// TIA Portal V20 export
// export: Created 2026-10-20T12:47:21.9915101Z, ExportSetting WithDefaults, DisplayName Totally Integrated Automation Portal, DisplayVersion V20 Update 6, DisplayName TIA Portal Openness, DisplayVersion V20 Update 6, DisplayName TIA Portal Version Control Interface, DisplayVersion V20 Update 6, DisplayName SINAMICS Startdrive Advanced, DisplayVersion V20 SP1, DisplayName SINAMICS Startdrive G130, G150, S120, S150, SINAMICS MV, G220, S200, S210, DisplayVersion V20 SP1, DisplayName SINAMICS Startdrive G110M, G120, G120C, G120D, G120P, G115D, DisplayVersion V20 SP1, DisplayName STEP 7 Professional, DisplayVersion V20 Update 6, DisplayName STEP 7 Safety, DisplayVersion V20 Update 2, DisplayName WinCC Basic/Comfort/Advanced, DisplayVersion V20 Update 6, DisplayName WinCC Unified, DisplayVersion V20 Update 6
FUNCTION "INPUTS" : Void   // FC25, SCL
{ S7_Optimized_Access := 'TRUE' }
VERSION : 0.1
// stored: AutoNumber true, IsIECCheckEnabled false, SetENOAutomatically false, UDAEnableTagReadback false
BEGIN
   REGION SYSTEM 1
       REGION EXTRACTOR CONVEYOR
           "Control_DB".ECnv_Sys[1].Inputs.Left := "CVTD1 SENSOR CONVEYOR LEFT";
           "Control_DB".ECnv_Sys[1].Inputs.Lpd1 := "CVTD1 SENSOR CONVEYOR LEFT (PALLET DETECT 1)";
           "Control_DB".ECnv_Sys[1].Inputs.Center := "CVTD1 SENSOR CONVEYOR CENTER";
           "Control_DB".ECnv_Sys[1].Inputs.Right := "CVTD1 SENSOR CONVEYOR RIGHT";
           "Control_DB".ECnv_Sys[1].Inputs.Rpd1 := "CVTD1 SENSOR CONVEYOR RIGHT (PALLET DETECT 1)";

           "T_OH_Left_1".TOF(IN := "CVTD1 OVERHANG LEFT" OR NOT "Control_DB".VTD_Sys[1].Running,
                             PT := T#200ms);
           "Control_DB".ECnv_Sys[1].Inputs.Overhang_Left := "T_OH_Left_1".Q;

           "T_OH_Right_1".TOF(IN := "CVTD1 OVERHANG RIGHT" OR NOT "Control_DB".VTD_Sys[1].Running,
                              PT := T#200ms);
           "Control_DB".ECnv_Sys[1].Inputs.Overhang_Right := "T_OH_Right_1".Q;

           "Control_DB".ECnv_Sys[1].Inputs.VFD_Status := "CVTD1_StatusWord";
           "Control_DB".ECnv_Sys[1].Inputs.VFD_ActualCurrent := WORD_TO_INT("CVTD1_ActualCurrent");
           "Control_DB".ECnv_Sys[1].Inputs.VFD_Speed_Actual := WORD_TO_INT("CVTD1_ActualSpeed");
           "Control_DB".ECnv_Sys[1].Inputs.VFD_ActualTorque := WORD_TO_INT("CVTD1_ActualTorque");
       END_REGION

       REGION BUFFER CONVEYORS
           REGION LEVEL 1
               //BUFFER CONVEYOR LEVEL 1 - CONVEYOR 1
               "Control_DB".LCnv_Sys[1].Cnv_Level[1].Cnv1.Inputs.Left := NOT "C1101 - SENSOR CNV LEFT";
               "Control_DB".LCnv_Sys[1].Cnv_Level[1].Cnv1.Inputs.Lpd1 := NOT "C1101 - SENSOR CNV LEFT (PALLET DETECT 1)";
               "Control_DB".LCnv_Sys[1].Cnv_Level[1].Cnv1.Inputs.Lpd2 := "C1101 - SENSOR CNV LEFT (PALLET DETECT 2)";
               "Control_DB".LCnv_Sys[1].Cnv_Level[1].Cnv1.Inputs.Right := NOT "C1101 - SENSOR CNV RIGHT";
               "Control_DB".LCnv_Sys[1].Cnv_Level[1].Cnv1.Inputs.Rpd1 := NOT "C1101 - SENSOR CNV RIGHT (PALLET DETECT 1)";
               "Control_DB".LCnv_Sys[1].Cnv_Level[1].Cnv1.Inputs.Rpd2 := NOT "C1101 - SENSOR CNV RIGHT (PALLET DETECT 2)";
               "Control_DB".LCnv_Sys[1].Cnv_Level[1].Cnv1.Inputs.Sdetect1 := NOT "C1101 - SHUTTLE IN POSITION 1";
               "Control_DB".LCnv_Sys[1].Cnv_Level[1].Cnv1.Inputs.Sdetect2 := NOT "C1101 - SHUTTLE IN POSITION 2";

               "Control_DB".LCnv_Sys[1].Cnv_Level[1].Cnv1.Inputs.VFD_Status := "C1101_StatusWord";
               "Control_DB".LCnv_Sys[1].Cnv_Level[1].Cnv1.Inputs.VFD_ActualCurrent := WORD_TO_INT("C1101_ActualCurrent");
               "Control_DB".LCnv_Sys[1].Cnv_Level[1].Cnv1.Inputs.VFD_Speed_Actual := WORD_TO_INT("C1101_ActualSpeed");
               "Control_DB".LCnv_Sys[1].Cnv_Level[1].Cnv1.Inputs.VFD_ActualTorque := WORD_TO_INT("C1101_ActualTorque");

               //BUFFER CONVEYOR LEVEL 1 - CONVEYOR 2
               "Control_DB".LCnv_Sys[1].Cnv_Level[1].Cnv2.Inputs.Left := NOT "C1201 - SENSOR CNV LEFT";
               "Control_DB".LCnv_Sys[1].Cnv_Level[1].Cnv2.Inputs.Lpd1 := NOT "C1201 - SENSOR CNV LEFT (PALLET DETECT 1)";
               "Control_DB".LCnv_Sys[1].Cnv_Level[1].Cnv2.Inputs.Lpd2 := NOT "C1201 - SENSOR CNV LEFT (PALLET DETECT 2)";
               "Control_DB".LCnv_Sys[1].Cnv_Level[1].Cnv2.Inputs.Right := NOT "C1201 - SENSOR CNV RIGHT";
               "Control_DB".LCnv_Sys[1].Cnv_Level[1].Cnv2.Inputs.Rpd1 := NOT "C1201 - SENSOR CNV RIGHT (PALLET DETECT 1)";
               "Control_DB".LCnv_Sys[1].Cnv_Level[1].Cnv2.Inputs.Rpd2 := NOT "C1201 - SENSOR CNV RIGHT (PALLET DETECT 2)";
               "Control_DB".LCnv_Sys[1].Cnv_Level[1].Cnv2.Inputs.Sdetect1 := NOT "C1201 - SHUTTLE IN POSITION 1";
               "Control_DB".LCnv_Sys[1].Cnv_Level[1].Cnv2.Inputs.Sdetect2 := NOT "C1201 - SHUTTLE IN POSITION 2";

               "Control_DB".LCnv_Sys[1].Cnv_Level[1].Cnv2.Inputs.VFD_Status := "C1201_StatusWord";
               "Control_DB".LCnv_Sys[1].Cnv_Level[1].Cnv2.Inputs.VFD_ActualCurrent := WORD_TO_INT("C1201_ActualCurrent");
               "Control_DB".LCnv_Sys[1].Cnv_Level[1].Cnv2.Inputs.VFD_Speed_Actual := WORD_TO_INT("C1201_ActualSpeed");
               "Control_DB".LCnv_Sys[1].Cnv_Level[1].Cnv2.Inputs.VFD_ActualTorque := WORD_TO_INT("C1201_ActualTorque");
           END_REGION

           REGION LEVEL 2
               //BUFFER CONVEYOR LEVEL 2 - CONVEYOR 1
               "Control_DB".LCnv_Sys[1].Cnv_Level[2].Cnv1.Inputs.Left := NOT "C1102 - SENSOR CNV LEFT";
               "Control_DB".LCnv_Sys[1].Cnv_Level[2].Cnv1.Inputs.Lpd1 := NOT "C1102 - SENSOR CNV LEFT (PALLET DETECT 1)";
               "Control_DB".LCnv_Sys[1].Cnv_Level[2].Cnv1.Inputs.Lpd2 := NOT "C1102 - SENSOR CNV LEFT (PALLET DETECT 2)";
               "Control_DB".LCnv_Sys[1].Cnv_Level[2].Cnv1.Inputs.Right := NOT "C1102 - SENSOR CNV RIGHT";
               "Control_DB".LCnv_Sys[1].Cnv_Level[2].Cnv1.Inputs.Rpd1 := NOT "C1102 - SENSOR CNV RIGHT (PALLET DETECT 1)";
               "Control_DB".LCnv_Sys[1].Cnv_Level[2].Cnv1.Inputs.Rpd2 := NOT "C1102 - SENSOR CNV RIGHT (PALLET DETECT 2)";
               "Control_DB".LCnv_Sys[1].Cnv_Level[2].Cnv1.Inputs.Sdetect1 := NOT "C1102 - SHUTTLE IN POSITION 1";
               "Control_DB".LCnv_Sys[1].Cnv_Level[2].Cnv1.Inputs.Sdetect2 := NOT "C1102 - SHUTTLE IN POSITION 2";
               "Control_DB".LCnv_Sys[1].Cnv_Level[2].Cnv1.Safety_Stop_Cnrl.Inputs.DP_Extended := "C1102 - SENSOR SAFETY PIN1 UP";
               "Control_DB".LCnv_Sys[1].Cnv_Level[2].Cnv1.Safety_Stop_Cnrl.Inputs.DP_Retracted := "C1102 - SENSOR SAFETY PIN1 DOWN";

               IF "Shuttle_MQTT_DB".Shuttle_MQTT[3].Message.Shuttle_Status.Position_ID = "Settings_DB".LCnv_Sys[1].Cnv_Level[2].Cnv1.Barcode_ID THEN
                   "Control_DB".LCnv_Sys[1].Cnv_Level[2].Cnv1.Inputs.Shuttle_High := "Shuttle_MQTT_DB".Shuttle_MQTT[3].Message.Shuttle_Status.Sensor_Inputs.%X13;
               ELSIF "Shuttle_MQTT_DB".Shuttle_MQTT[4].Message.Shuttle_Status.Position_ID = "Settings_DB".LCnv_Sys[1].Cnv_Level[2].Cnv1.Barcode_ID THEN
                   "Control_DB".LCnv_Sys[1].Cnv_Level[2].Cnv1.Inputs.Shuttle_High := "Shuttle_MQTT_DB".Shuttle_MQTT[4].Message.Shuttle_Status.Sensor_Inputs.%X13;
               ELSIF "Shuttle_MQTT_DB".Shuttle_MQTT[5].Message.Shuttle_Status.Position_ID = "Settings_DB".LCnv_Sys[1].Cnv_Level[2].Cnv1.Barcode_ID THEN
                   "Control_DB".LCnv_Sys[1].Cnv_Level[2].Cnv1.Inputs.Shuttle_High := "Shuttle_MQTT_DB".Shuttle_MQTT[5].Message.Shuttle_Status.Sensor_Inputs.%X13;
               END_IF;

               "Control_DB".LCnv_Sys[1].Cnv_Level[2].Cnv1.Inputs.VFD_Status := "C1102_StatusWord";
               "Control_DB".LCnv_Sys[1].Cnv_Level[2].Cnv1.Inputs.VFD_ActualCurrent := WORD_TO_INT("C1102_ActualCurrent");
               "Control_DB".LCnv_Sys[1].Cnv_Level[2].Cnv1.Inputs.VFD_Speed_Actual := WORD_TO_INT("C1102_ActualSpeed");
               "Control_DB".LCnv_Sys[1].Cnv_Level[2].Cnv1.Inputs.VFD_ActualTorque := "C1102_ActualTorque";

               //BUFFER CONVEYOR LEVEL 2 - CONVEYOR 2
               "Control_DB".LCnv_Sys[1].Cnv_Level[2].Cnv2.Inputs.Left := NOT "C1202 - SENSOR CNV LEFT";
               "Control_DB".LCnv_Sys[1].Cnv_Level[2].Cnv2.Inputs.Lpd1 := NOT "C1202 - SENSOR CNV LEFT (PALLET DETECT 1)";
               "Control_DB".LCnv_Sys[1].Cnv_Level[2].Cnv2.Inputs.Lpd2 := NOT "C1202 - SENSOR CNV LEFT (PALLET DETECT 2)";
               "Control_DB".LCnv_Sys[1].Cnv_Level[2].Cnv2.Inputs.Right := NOT "C1202 - SENSOR CNV RIGHT";
               "Control_DB".LCnv_Sys[1].Cnv_Level[2].Cnv2.Inputs.Rpd1 := NOT "C1202 - SENSOR CNV RIGHT (PALLET DETECT 1)";
               "Control_DB".LCnv_Sys[1].Cnv_Level[2].Cnv2.Inputs.Rpd2 := NOT "C1202 - SENSOR CNV RIGHT (PALLET DETECT 2)";
               "Control_DB".LCnv_Sys[1].Cnv_Level[2].Cnv2.Inputs.Sdetect1 := NOT "C1202 - SHUTTLE IN POSITION 1";
               "Control_DB".LCnv_Sys[1].Cnv_Level[2].Cnv2.Inputs.Sdetect2 := NOT "C1202 - SHUTTLE IN POSITION 2";
               "Control_DB".LCnv_Sys[1].Cnv_Level[2].Cnv2.Safety_Stop_Cnrl.Inputs.DP_Extended := "C1202 - SENSOR SAFETY PIN1 UP";
               "Control_DB".LCnv_Sys[1].Cnv_Level[2].Cnv2.Safety_Stop_Cnrl.Inputs.DP_Retracted := "C1202 - SENSOR SAFETY PIN1 DOWN";

               IF "Shuttle_MQTT_DB".Shuttle_MQTT[3].Message.Shuttle_Status.Position_ID = "Settings_DB".LCnv_Sys[1].Cnv_Level[2].Cnv2.Barcode_ID THEN
                   "Control_DB".LCnv_Sys[1].Cnv_Level[2].Cnv2.Inputs.Shuttle_High := "Shuttle_MQTT_DB".Shuttle_MQTT[3].Message.Shuttle_Status.Sensor_Inputs.%X13;
               ELSIF "Shuttle_MQTT_DB".Shuttle_MQTT[4].Message.Shuttle_Status.Position_ID = "Settings_DB".LCnv_Sys[1].Cnv_Level[2].Cnv2.Barcode_ID THEN
                   "Control_DB".LCnv_Sys[1].Cnv_Level[2].Cnv2.Inputs.Shuttle_High := "Shuttle_MQTT_DB".Shuttle_MQTT[4].Message.Shuttle_Status.Sensor_Inputs.%X13;
               ELSIF "Shuttle_MQTT_DB".Shuttle_MQTT[5].Message.Shuttle_Status.Position_ID = "Settings_DB".LCnv_Sys[1].Cnv_Level[2].Cnv2.Barcode_ID THEN
                   "Control_DB".LCnv_Sys[1].Cnv_Level[2].Cnv2.Inputs.Shuttle_High := "Shuttle_MQTT_DB".Shuttle_MQTT[5].Message.Shuttle_Status.Sensor_Inputs.%X13;
               END_IF;

               "Control_DB".LCnv_Sys[1].Cnv_Level[2].Cnv2.Inputs.VFD_Status := "C1202_StatusWord";
               "Control_DB".LCnv_Sys[1].Cnv_Level[2].Cnv2.Inputs.VFD_ActualCurrent := WORD_TO_INT("C1202_ActualCurrent");
               "Control_DB".LCnv_Sys[1].Cnv_Level[2].Cnv2.Inputs.VFD_Speed_Actual := WORD_TO_INT("C1202_ActualSpeed");
               "Control_DB".LCnv_Sys[1].Cnv_Level[2].Cnv2.Inputs.VFD_ActualTorque := "C1202_ActualTorque";
           END_REGION

           REGION LEVEL 3
               //BUFFER CONVEYOR LEVEL 3 - CONVEYOR 1
               "Control_DB".LCnv_Sys[1].Cnv_Level[3].Cnv1.Inputs.Left := NOT "C1103 - SENSOR CNV LEFT";
               "Control_DB".LCnv_Sys[1].Cnv_Level[3].Cnv1.Inputs.Lpd1 := NOT "C1103 - SENSOR CNV LEFT (PALLET DETECT 1)";
               "Control_DB".LCnv_Sys[1].Cnv_Level[3].Cnv1.Inputs.Lpd2 := NOT "C1103 - SENSOR CNV LEFT (PALLET DETECT 2)";
               "Control_DB".LCnv_Sys[1].Cnv_Level[3].Cnv1.Inputs.Right := NOT "C1103 - SENSOR CNV RIGHT";
               "Control_DB".LCnv_Sys[1].Cnv_Level[3].Cnv1.Inputs.Rpd1 := NOT "C1103 - SENSOR CNV RIGHT (PALLET DETECT 1)";
               "Control_DB".LCnv_Sys[1].Cnv_Level[3].Cnv1.Inputs.Rpd2 := NOT "C1103 - SENSOR CNV RIGHT (PALLET DETECT 2)";
               "Control_DB".LCnv_Sys[1].Cnv_Level[3].Cnv1.Inputs.Sdetect1 := NOT "C1103 - SHUTTLE IN POSITION 1";
               "Control_DB".LCnv_Sys[1].Cnv_Level[3].Cnv1.Inputs.Sdetect2 := NOT "C1103 - SHUTTLE IN POSITION 2";
               "Control_DB".LCnv_Sys[1].Cnv_Level[3].Cnv1.Safety_Stop_Cnrl.Inputs.DP_Extended := "C1103 - SENSOR SAFETY PIN1 UP";
               "Control_DB".LCnv_Sys[1].Cnv_Level[3].Cnv1.Safety_Stop_Cnrl.Inputs.DP_Retracted := "C1103 - SENSOR SAFETY PIN1 DOWN";

               "Control_DB".LCnv_Sys[1].Cnv_Level[3].Cnv1.Inputs.VFD_Status := "C1103_StatusWord";
               "Control_DB".LCnv_Sys[1].Cnv_Level[3].Cnv1.Inputs.VFD_ActualCurrent := WORD_TO_INT("C1103_ActualCurrent");
               "Control_DB".LCnv_Sys[1].Cnv_Level[3].Cnv1.Inputs.VFD_Speed_Actual := WORD_TO_INT("C1103_ActualSpeed");
               "Control_DB".LCnv_Sys[1].Cnv_Level[3].Cnv1.Inputs.VFD_ActualTorque := "C1103_ActualTorque";

               //BUFFER CONVEYOR LEVEL 3 - CONVEYOR 2
               "Control_DB".LCnv_Sys[1].Cnv_Level[3].Cnv2.Inputs.Left := NOT "C1203 - SENSOR CNV LEFT";
               "Control_DB".LCnv_Sys[1].Cnv_Level[3].Cnv2.Inputs.Lpd1 := NOT "C1203 - SENSOR CNV LEFT (PALLET DETECT 1)";
               "Control_DB".LCnv_Sys[1].Cnv_Level[3].Cnv2.Inputs.Lpd2 := NOT "C1203 - SENSOR CNV LEFT (PALLET DETECT 2)";
               "Control_DB".LCnv_Sys[1].Cnv_Level[3].Cnv2.Inputs.Right := NOT "C1203 - SENSOR CNV RIGHT";
               "Control_DB".LCnv_Sys[1].Cnv_Level[3].Cnv2.Inputs.Rpd1 := NOT "C1203 - SENSOR CNV RIGHT (PALLET DETECT 1)";
               "Control_DB".LCnv_Sys[1].Cnv_Level[3].Cnv2.Inputs.Rpd2 := NOT "C1203 - SENSOR CNV RIGHT (PALLET DETECT 2)";
               "Control_DB".LCnv_Sys[1].Cnv_Level[3].Cnv2.Inputs.Sdetect1 := NOT "C1203 - SHUTTLE IN POSITION 1";
               "Control_DB".LCnv_Sys[1].Cnv_Level[3].Cnv2.Inputs.Sdetect2 := NOT "C1203 - SHUTTLE IN POSITION 2";
               "Control_DB".LCnv_Sys[1].Cnv_Level[3].Cnv2.Safety_Stop_Cnrl.Inputs.DP_Extended := "C1203 - SENSOR SAFETY PIN1 UP";
               "Control_DB".LCnv_Sys[1].Cnv_Level[3].Cnv2.Safety_Stop_Cnrl.Inputs.DP_Retracted := "C1203 - SENSOR SAFETY PIN1 DOWN";

               "Control_DB".LCnv_Sys[1].Cnv_Level[3].Cnv2.Inputs.VFD_Status := "C1203_StatusWord";
               "Control_DB".LCnv_Sys[1].Cnv_Level[3].Cnv2.Inputs.VFD_ActualCurrent := WORD_TO_INT("C1203_ActualCurrent");
               "Control_DB".LCnv_Sys[1].Cnv_Level[3].Cnv2.Inputs.VFD_Speed_Actual := WORD_TO_INT("C1203_ActualSpeed");
               "Control_DB".LCnv_Sys[1].Cnv_Level[3].Cnv2.Inputs.VFD_ActualTorque := "C1203_ActualTorque";
           END_REGION

           REGION LEVEL 4
               //BUFFER CONVEYOR LEVEL 4 - CONVEYOR 1
               "Control_DB".LCnv_Sys[1].Cnv_Level[4].Cnv1.Inputs.Left := NOT "C1104 - SENSOR CNV LEFT";
               "Control_DB".LCnv_Sys[1].Cnv_Level[4].Cnv1.Inputs.Lpd1 := NOT "C1104 - SENSOR CNV LEFT (PALLET DETECT 1)";
               "Control_DB".LCnv_Sys[1].Cnv_Level[4].Cnv1.Inputs.Lpd2 := NOT "C1104 - SENSOR CNV LEFT (PALLET DETECT 2)";
               "Control_DB".LCnv_Sys[1].Cnv_Level[4].Cnv1.Inputs.Right := NOT "C1104 - SENSOR CNV RIGHT";
               "Control_DB".LCnv_Sys[1].Cnv_Level[4].Cnv1.Inputs.Rpd1 := NOT "C1104 - SENSOR CNV RIGHT (PALLET DETECT 1)";
               "Control_DB".LCnv_Sys[1].Cnv_Level[4].Cnv1.Inputs.Rpd2 := NOT "C1104 - SENSOR CNV RIGHT (PALLET DETECT 2)";
               "Control_DB".LCnv_Sys[1].Cnv_Level[4].Cnv1.Inputs.Sdetect1 := NOT "C1104 - SHUTTLE IN POSITION 1";
               "Control_DB".LCnv_Sys[1].Cnv_Level[4].Cnv1.Inputs.Sdetect2 := NOT "C1104 - SHUTTLE IN POSITION 2";
               "Control_DB".LCnv_Sys[1].Cnv_Level[4].Cnv1.Safety_Stop_Cnrl.Inputs.DP_Extended := "C1104 - SENSOR SAFETY PIN1 UP";
               "Control_DB".LCnv_Sys[1].Cnv_Level[4].Cnv1.Safety_Stop_Cnrl.Inputs.DP_Retracted := "C1104 - SENSOR SAFETY PIN1 DOWN";

               "Control_DB".LCnv_Sys[1].Cnv_Level[4].Cnv1.Inputs.VFD_Status := "C1104_StatusWord";
               "Control_DB".LCnv_Sys[1].Cnv_Level[4].Cnv1.Inputs.VFD_ActualCurrent := WORD_TO_INT("C1104_ActualCurrent");
               "Control_DB".LCnv_Sys[1].Cnv_Level[4].Cnv1.Inputs.VFD_Speed_Actual := WORD_TO_INT("C1104_ActualSpeed");
               "Control_DB".LCnv_Sys[1].Cnv_Level[4].Cnv1.Inputs.VFD_ActualTorque := "C1104_ActualTorque";

               //BUFFER CONVEYOR LEVEL 4 - CONVEYOR 2
               "Control_DB".LCnv_Sys[1].Cnv_Level[4].Cnv2.Inputs.Left := NOT "C1204 - SENSOR CNV LEFT";
               "Control_DB".LCnv_Sys[1].Cnv_Level[4].Cnv2.Inputs.Lpd1 := NOT "C1204 - SENSOR CNV LEFT (PALLET DETECT 1)";
               "Control_DB".LCnv_Sys[1].Cnv_Level[4].Cnv2.Inputs.Lpd2 := NOT "C1204 - SENSOR CNV LEFT (PALLET DETECT 2)";
               "Control_DB".LCnv_Sys[1].Cnv_Level[4].Cnv2.Inputs.Right := NOT "C1204 - SENSOR CNV RIGHT";
               "Control_DB".LCnv_Sys[1].Cnv_Level[4].Cnv2.Inputs.Rpd1 := NOT "C1204 - SENSOR CNV RIGHT (PALLET DETECT 1)";
               "Control_DB".LCnv_Sys[1].Cnv_Level[4].Cnv2.Inputs.Rpd2 := NOT "C1204 - SENSOR CNV RIGHT (PALLET DETECT 2)";
               "Control_DB".LCnv_Sys[1].Cnv_Level[4].Cnv2.Inputs.Sdetect1 := NOT "C1204 - SHUTTLE IN POSITION 1";
               "Control_DB".LCnv_Sys[1].Cnv_Level[4].Cnv2.Inputs.Sdetect2 := NOT "C1204 - SHUTTLE IN POSITION 2";
               "Control_DB".LCnv_Sys[1].Cnv_Level[4].Cnv2.Safety_Stop_Cnrl.Inputs.DP_Extended := "C1204 - SENSOR SAFETY PIN1 UP";
               "Control_DB".LCnv_Sys[1].Cnv_Level[4].Cnv2.Safety_Stop_Cnrl.Inputs.DP_Retracted := "C1204 - SENSOR SAFETY PIN1 DOWN";

               "Control_DB".LCnv_Sys[1].Cnv_Level[4].Cnv2.Inputs.VFD_Status := "C1204_StatusWord";
               "Control_DB".LCnv_Sys[1].Cnv_Level[4].Cnv2.Inputs.VFD_ActualCurrent := WORD_TO_INT("C1204_ActualCurrent");
               "Control_DB".LCnv_Sys[1].Cnv_Level[4].Cnv2.Inputs.VFD_Speed_Actual := WORD_TO_INT("C1204_ActualSpeed");
               "Control_DB".LCnv_Sys[1].Cnv_Level[4].Cnv2.Inputs.VFD_ActualTorque := "C1204_ActualTorque";
           END_REGION

           REGION LEVEL 5
               //BUFFER CONVEYOR LEVEL 5 - CONVEYOR 1
               "Control_DB".LCnv_Sys[1].Cnv_Level[5].Cnv1.Inputs.Left := NOT "C1105 - SENSOR CNV LEFT";
               "Control_DB".LCnv_Sys[1].Cnv_Level[5].Cnv1.Inputs.Lpd1 := NOT "C1105 - SENSOR CNV LEFT (PALLET DETECT 1)";
               "Control_DB".LCnv_Sys[1].Cnv_Level[5].Cnv1.Inputs.Lpd2 := NOT "C1105 - SENSOR CNV LEFT (PALLET DETECT 2)";
               "Control_DB".LCnv_Sys[1].Cnv_Level[5].Cnv1.Inputs.Right := NOT "C1105 - SENSOR CNV RIGHT";
               "Control_DB".LCnv_Sys[1].Cnv_Level[5].Cnv1.Inputs.Rpd1 := NOT "C1105 - SENSOR CNV RIGHT (PALLET DETECT 1)";
               "Control_DB".LCnv_Sys[1].Cnv_Level[5].Cnv1.Inputs.Rpd2 := NOT "C1105 - SENSOR CNV RIGHT (PALLET DETECT 2)";
               "Control_DB".LCnv_Sys[1].Cnv_Level[5].Cnv1.Inputs.Sdetect1 := NOT "C1105 - SHUTTLE IN POSITION 1";
               "Control_DB".LCnv_Sys[1].Cnv_Level[5].Cnv1.Inputs.Sdetect2 := NOT "C1105 - SHUTTLE IN POSITION 2";
               "Control_DB".LCnv_Sys[1].Cnv_Level[5].Cnv1.Safety_Stop_Cnrl.Inputs.DP_Extended := "C1105 - SENSOR SAFETY PIN1 UP";
               "Control_DB".LCnv_Sys[1].Cnv_Level[5].Cnv1.Safety_Stop_Cnrl.Inputs.DP_Retracted := "C1105 - SENSOR SAFETY PIN1 DOWN";

               "Control_DB".LCnv_Sys[1].Cnv_Level[5].Cnv1.Inputs.VFD_Status := "C1105_StatusWord";
               "Control_DB".LCnv_Sys[1].Cnv_Level[5].Cnv1.Inputs.VFD_ActualCurrent := WORD_TO_INT("C1105_ActualCurrent");
               "Control_DB".LCnv_Sys[1].Cnv_Level[5].Cnv1.Inputs.VFD_Speed_Actual := WORD_TO_INT("C1105_ActualSpeed");
               "Control_DB".LCnv_Sys[1].Cnv_Level[5].Cnv1.Inputs.VFD_ActualTorque := "C1105_ActualTorque";

               //BUFFER CONVEYOR LEVEL 5 - CONVEYOR 2
               "Control_DB".LCnv_Sys[1].Cnv_Level[5].Cnv2.Inputs.Left := NOT "C1205 - SENSOR CNV LEFT";
               "Control_DB".LCnv_Sys[1].Cnv_Level[5].Cnv2.Inputs.Lpd1 := NOT "C1205 - SENSOR CNV LEFT (PALLET DETECT 1)";
               "Control_DB".LCnv_Sys[1].Cnv_Level[5].Cnv2.Inputs.Lpd2 := NOT "C1205 - SENSOR CNV LEFT (PALLET DETECT 2)";
               "Control_DB".LCnv_Sys[1].Cnv_Level[5].Cnv2.Inputs.Right := NOT "C1205 - SENSOR CNV RIGHT";
               "Control_DB".LCnv_Sys[1].Cnv_Level[5].Cnv2.Inputs.Rpd1 := NOT "C1205 - SENSOR CNV RIGHT (PALLET DETECT 1)";
               "Control_DB".LCnv_Sys[1].Cnv_Level[5].Cnv2.Inputs.Rpd2 := NOT "C1205 - SENSOR CNV RIGHT (PALLET DETECT 2)";
               "Control_DB".LCnv_Sys[1].Cnv_Level[5].Cnv2.Inputs.Sdetect1 := NOT "C1205 - SHUTTLE IN POSITION 1";
               "Control_DB".LCnv_Sys[1].Cnv_Level[5].Cnv2.Inputs.Sdetect2 := NOT "C1205 - SHUTTLE IN POSITION 2";
               "Control_DB".LCnv_Sys[1].Cnv_Level[5].Cnv2.Safety_Stop_Cnrl.Inputs.DP_Extended := "C1205 - SENSOR SAFETY PIN1 UP";
               "Control_DB".LCnv_Sys[1].Cnv_Level[5].Cnv2.Safety_Stop_Cnrl.Inputs.DP_Retracted := "C1205 - SENSOR SAFETY PIN1 DOWN";

               "Control_DB".LCnv_Sys[1].Cnv_Level[5].Cnv2.Inputs.VFD_Status := "C1205_StatusWord";
               "Control_DB".LCnv_Sys[1].Cnv_Level[5].Cnv2.Inputs.VFD_ActualCurrent := WORD_TO_INT("C1205_ActualCurrent");
               "Control_DB".LCnv_Sys[1].Cnv_Level[5].Cnv2.Inputs.VFD_Speed_Actual := WORD_TO_INT("C1205_ActualSpeed");
               "Control_DB".LCnv_Sys[1].Cnv_Level[5].Cnv2.Inputs.VFD_ActualTorque := "C1205_ActualTorque";
           END_REGION

           REGION LEVEL 6
               //BUFFER CONVEYOR LEVEL 6 - CONVEYOR 1
               "Control_DB".LCnv_Sys[1].Cnv_Level[6].Cnv1.Inputs.Left := NOT "C1106 - SENSOR CNV LEFT";
               "Control_DB".LCnv_Sys[1].Cnv_Level[6].Cnv1.Inputs.Lpd1 := NOT "C1106 - SENSOR CNV LEFT (PALLET DETECT 1)";
               "Control_DB".LCnv_Sys[1].Cnv_Level[6].Cnv1.Inputs.Lpd2 := NOT "C1106 - SENSOR CNV LEFT (PALLET DETECT 2)";
               "Control_DB".LCnv_Sys[1].Cnv_Level[6].Cnv1.Inputs.Right := NOT "C1106 - SENSOR CNV RIGHT";
               "Control_DB".LCnv_Sys[1].Cnv_Level[6].Cnv1.Inputs.Rpd1 := NOT "C1106 - SENSOR CNV RIGHT (PALLET DETECT 1)";
               "Control_DB".LCnv_Sys[1].Cnv_Level[6].Cnv1.Inputs.Rpd2 := NOT "C1106 - SENSOR CNV RIGHT (PALLET DETECT 2)";
               "Control_DB".LCnv_Sys[1].Cnv_Level[6].Cnv1.Inputs.Sdetect1 := NOT "C1106 - SHUTTLE IN POSITION 1";
               "Control_DB".LCnv_Sys[1].Cnv_Level[6].Cnv1.Inputs.Sdetect2 := NOT "C1106 - SHUTTLE IN POSITION 2";
               "Control_DB".LCnv_Sys[1].Cnv_Level[6].Cnv1.Safety_Stop_Cnrl.Inputs.DP_Extended := "C1106 - SENSOR SAFETY PIN1 UP";
               "Control_DB".LCnv_Sys[1].Cnv_Level[6].Cnv1.Safety_Stop_Cnrl.Inputs.DP_Retracted := "C1106 - SENSOR SAFETY PIN1 DOWN";

               "Control_DB".LCnv_Sys[1].Cnv_Level[6].Cnv1.Inputs.VFD_Status := "C1106_StatusWord";
               "Control_DB".LCnv_Sys[1].Cnv_Level[6].Cnv1.Inputs.VFD_ActualCurrent := WORD_TO_INT("C1106_ActualCurrent");
               "Control_DB".LCnv_Sys[1].Cnv_Level[6].Cnv1.Inputs.VFD_Speed_Actual := WORD_TO_INT("C1106_ActualSpeed");
               "Control_DB".LCnv_Sys[1].Cnv_Level[6].Cnv1.Inputs.VFD_ActualTorque := "C1106_ActualTorque";

               //BUFFER CONVEYOR LEVEL 6 - CONVEYOR 2
               "Control_DB".LCnv_Sys[1].Cnv_Level[6].Cnv2.Inputs.Left := NOT "C1206 - SENSOR CNV LEFT";
               "Control_DB".LCnv_Sys[1].Cnv_Level[6].Cnv2.Inputs.Lpd1 := NOT "C1206 - SENSOR CNV LEFT (PALLET DETECT 1)";
               "Control_DB".LCnv_Sys[1].Cnv_Level[6].Cnv2.Inputs.Lpd2 := NOT "C1206 - SENSOR CNV LEFT (PALLET DETECT 2)";
               "Control_DB".LCnv_Sys[1].Cnv_Level[6].Cnv2.Inputs.Right := NOT "C1206 - SENSOR CNV RIGHT";
               "Control_DB".LCnv_Sys[1].Cnv_Level[6].Cnv2.Inputs.Rpd1 := NOT "C1206 - SENSOR CNV RIGHT (PALLET DETECT 1)";
               "Control_DB".LCnv_Sys[1].Cnv_Level[6].Cnv2.Inputs.Rpd2 := NOT "C1206 - SENSOR CNV RIGHT (PALLET DETECT 2)";
               "Control_DB".LCnv_Sys[1].Cnv_Level[6].Cnv2.Inputs.Sdetect1 := NOT "C1206 - SHUTTLE IN POSITION 1";
               "Control_DB".LCnv_Sys[1].Cnv_Level[6].Cnv2.Inputs.Sdetect2 := NOT "C1206 - SHUTTLE IN POSITION 2";
               "Control_DB".LCnv_Sys[1].Cnv_Level[6].Cnv2.Safety_Stop_Cnrl.Inputs.DP_Extended := "C1206 - SENSOR SAFETY PIN1 UP";
               "Control_DB".LCnv_Sys[1].Cnv_Level[6].Cnv2.Safety_Stop_Cnrl.Inputs.DP_Retracted := "C1206 - SENSOR SAFETY PIN1 DOWN";

               "Control_DB".LCnv_Sys[1].Cnv_Level[6].Cnv2.Inputs.VFD_Status := "C1206_StatusWord";
               "Control_DB".LCnv_Sys[1].Cnv_Level[6].Cnv2.Inputs.VFD_ActualCurrent := WORD_TO_INT("C1206_ActualCurrent");
               "Control_DB".LCnv_Sys[1].Cnv_Level[6].Cnv2.Inputs.VFD_Speed_Actual := WORD_TO_INT("C1206_ActualSpeed");
               "Control_DB".LCnv_Sys[1].Cnv_Level[6].Cnv2.Inputs.VFD_ActualTorque := "C1206_ActualTorque";
           END_REGION

           REGION LEVEL 7
               //BUFFER CONVEYOR LEVEL 7 - CONVEYOR 1
               "Control_DB".LCnv_Sys[1].Cnv_Level[7].Cnv1.Inputs.Left := NOT "C1107 - SENSOR CNV LEFT";
               "Control_DB".LCnv_Sys[1].Cnv_Level[7].Cnv1.Inputs.Lpd1 := NOT "C1107 - SENSOR CNV LEFT (PALLET DETECT 1)";
               "Control_DB".LCnv_Sys[1].Cnv_Level[7].Cnv1.Inputs.Lpd2 := NOT "C1107 - SENSOR CNV LEFT (PALLET DETECT 2)";
               "Control_DB".LCnv_Sys[1].Cnv_Level[7].Cnv1.Inputs.Right := NOT "C1107 - SENSOR CNV RIGHT";
               "Control_DB".LCnv_Sys[1].Cnv_Level[7].Cnv1.Inputs.Rpd1 := NOT "C1107 - SENSOR CNV RIGHT (PALLET DETECT 1)";
               "Control_DB".LCnv_Sys[1].Cnv_Level[7].Cnv1.Inputs.Rpd2 := NOT "C1107 - SENSOR CNV RIGHT (PALLET DETECT 2)";
               "Control_DB".LCnv_Sys[1].Cnv_Level[7].Cnv1.Inputs.Sdetect1 := NOT "C1107 - SHUTTLE IN POSITION 1";
               "Control_DB".LCnv_Sys[1].Cnv_Level[7].Cnv1.Inputs.Sdetect2 := NOT "C1107 - SHUTTLE IN POSITION 2";
               "Control_DB".LCnv_Sys[1].Cnv_Level[7].Cnv1.Safety_Stop_Cnrl.Inputs.DP_Extended := "C1107 - SENSOR SAFETY PIN1 UP";
               "Control_DB".LCnv_Sys[1].Cnv_Level[7].Cnv1.Safety_Stop_Cnrl.Inputs.DP_Retracted := "C1107 - SENSOR SAFETY PIN1 DOWN";

               "Control_DB".LCnv_Sys[1].Cnv_Level[7].Cnv1.Inputs.VFD_Status := "C1107_StatusWord";
               "Control_DB".LCnv_Sys[1].Cnv_Level[7].Cnv1.Inputs.VFD_ActualCurrent := WORD_TO_INT("C1107_ActualCurrent");
               "Control_DB".LCnv_Sys[1].Cnv_Level[7].Cnv1.Inputs.VFD_Speed_Actual := WORD_TO_INT("C1107_ActualSpeed");
               "Control_DB".LCnv_Sys[1].Cnv_Level[7].Cnv1.Inputs.VFD_ActualTorque := "C1107_ActualTorque";

               //BUFFER CONVEYOR LEVEL 7 - CONVEYOR 2
               "Control_DB".LCnv_Sys[1].Cnv_Level[7].Cnv2.Inputs.Left := NOT "C1207 - SENSOR CNV LEFT";
               "Control_DB".LCnv_Sys[1].Cnv_Level[7].Cnv2.Inputs.Lpd1 := NOT "C1207 - SENSOR CNV LEFT (PALLET DETECT 1)";
               "Control_DB".LCnv_Sys[1].Cnv_Level[7].Cnv2.Inputs.Lpd2 := NOT "C1207 - SENSOR CNV LEFT (PALLET DETECT 2)";
               "Control_DB".LCnv_Sys[1].Cnv_Level[7].Cnv2.Inputs.Right := NOT "C1207 - SENSOR CNV RIGHT";
               "Control_DB".LCnv_Sys[1].Cnv_Level[7].Cnv2.Inputs.Rpd1 := NOT "C1207 - SENSOR CNV RIGHT (PALLET DETECT 1)";
               "Control_DB".LCnv_Sys[1].Cnv_Level[7].Cnv2.Inputs.Rpd2 := NOT "C1207 - SENSOR CNV RIGHT (PALLET DETECT 2)";
               "Control_DB".LCnv_Sys[1].Cnv_Level[7].Cnv2.Inputs.Sdetect1 := NOT "C1207 - SHUTTLE IN POSITION 1";
               "Control_DB".LCnv_Sys[1].Cnv_Level[7].Cnv2.Inputs.Sdetect2 := NOT "C1207 - SHUTTLE IN POSITION 2";
               "Control_DB".LCnv_Sys[1].Cnv_Level[7].Cnv2.Safety_Stop_Cnrl.Inputs.DP_Extended := "C1207 - SENSOR SAFETY PIN1 UP";
               "Control_DB".LCnv_Sys[1].Cnv_Level[7].Cnv2.Safety_Stop_Cnrl.Inputs.DP_Retracted := "C1207 - SENSOR SAFETY PIN1 DOWN";

               "Control_DB".LCnv_Sys[1].Cnv_Level[7].Cnv2.Inputs.VFD_Status := "C1207_StatusWord";
               "Control_DB".LCnv_Sys[1].Cnv_Level[7].Cnv2.Inputs.VFD_ActualCurrent := WORD_TO_INT("C1207_ActualCurrent");
               "Control_DB".LCnv_Sys[1].Cnv_Level[7].Cnv2.Inputs.VFD_Speed_Actual := WORD_TO_INT("C1207_ActualSpeed");
               "Control_DB".LCnv_Sys[1].Cnv_Level[7].Cnv2.Inputs.VFD_ActualTorque := "C1207_ActualTorque";
           END_REGION

           REGION LEVEL 8
               //BUFFER CONVEYOR LEVEL 8 - CONVEYOR 1
               "Control_DB".LCnv_Sys[1].Cnv_Level[8].Cnv1.Inputs.Left := NOT "C1108 - SENSOR CNV LEFT";
               "Control_DB".LCnv_Sys[1].Cnv_Level[8].Cnv1.Inputs.Lpd1 := NOT "C1108 - SENSOR CNV LEFT (PALLET DETECT 1)";
               "Control_DB".LCnv_Sys[1].Cnv_Level[8].Cnv1.Inputs.Lpd2 := NOT "C1108 - SENSOR CNV LEFT (PALLET DETECT 2)";
               "Control_DB".LCnv_Sys[1].Cnv_Level[8].Cnv1.Inputs.Right := NOT "C1108 - SENSOR CNV RIGHT";
               "Control_DB".LCnv_Sys[1].Cnv_Level[8].Cnv1.Inputs.Rpd1 := NOT "C1108 - SENSOR CNV RIGHT (PALLET DETECT 1)";
               "Control_DB".LCnv_Sys[1].Cnv_Level[8].Cnv1.Inputs.Rpd2 := NOT "C1108 - SENSOR CNV RIGHT (PALLET DETECT 2)";
               "Control_DB".LCnv_Sys[1].Cnv_Level[8].Cnv1.Inputs.Sdetect1 := NOT "C1108 - SHUTTLE IN POSITION 1";
               "Control_DB".LCnv_Sys[1].Cnv_Level[8].Cnv1.Inputs.Sdetect2 := NOT "C1108 - SHUTTLE IN POSITION 2";
               "Control_DB".LCnv_Sys[1].Cnv_Level[8].Cnv1.Safety_Stop_Cnrl.Inputs.DP_Extended := "C1108 - SENSOR SAFETY PIN1 UP";
               "Control_DB".LCnv_Sys[1].Cnv_Level[8].Cnv1.Safety_Stop_Cnrl.Inputs.DP_Retracted := "C1108 - SENSOR SAFETY PIN1 DOWN";

               "Control_DB".LCnv_Sys[1].Cnv_Level[8].Cnv1.Inputs.VFD_Status := "C1108_StatusWord";
               "Control_DB".LCnv_Sys[1].Cnv_Level[8].Cnv1.Inputs.VFD_ActualCurrent := WORD_TO_INT("C1108_ActualCurrent");
               "Control_DB".LCnv_Sys[1].Cnv_Level[8].Cnv1.Inputs.VFD_Speed_Actual := WORD_TO_INT("C1108_ActualSpeed");
               "Control_DB".LCnv_Sys[1].Cnv_Level[8].Cnv1.Inputs.VFD_ActualTorque := "C1108_ActualTorque";

               //BUFFER CONVEYOR LEVEL 8 - CONVEYOR 2
               "Control_DB".LCnv_Sys[1].Cnv_Level[8].Cnv2.Inputs.Left := NOT "C1208 - SENSOR CNV LEFT";
               "Control_DB".LCnv_Sys[1].Cnv_Level[8].Cnv2.Inputs.Lpd1 := NOT "C1208 - SENSOR CNV LEFT (PALLET DETECT 1)";
               "Control_DB".LCnv_Sys[1].Cnv_Level[8].Cnv2.Inputs.Lpd2 := NOT "C1208 - SENSOR CNV LEFT (PALLET DETECT 2)";
               "Control_DB".LCnv_Sys[1].Cnv_Level[8].Cnv2.Inputs.Right := NOT "C1208 - SENSOR CNV RIGHT";
               "Control_DB".LCnv_Sys[1].Cnv_Level[8].Cnv2.Inputs.Rpd1 := NOT "C1208 - SENSOR CNV RIGHT (PALLET DETECT 1)";
               "Control_DB".LCnv_Sys[1].Cnv_Level[8].Cnv2.Inputs.Rpd2 := NOT "C1208 - SENSOR CNV RIGHT (PALLET DETECT 2)";
               "Control_DB".LCnv_Sys[1].Cnv_Level[8].Cnv2.Inputs.Sdetect1 := NOT "C1208 - SHUTTLE IN POSITION 1";
               "Control_DB".LCnv_Sys[1].Cnv_Level[8].Cnv2.Inputs.Sdetect2 := NOT "C1208 - SHUTTLE IN POSITION 2";
               "Control_DB".LCnv_Sys[1].Cnv_Level[8].Cnv2.Safety_Stop_Cnrl.Inputs.DP_Extended := "C1208 - SENSOR SAFETY PIN1 UP";
               "Control_DB".LCnv_Sys[1].Cnv_Level[8].Cnv2.Safety_Stop_Cnrl.Inputs.DP_Retracted := "C1208 - SENSOR SAFETY PIN1 DOWN";

               "Control_DB".LCnv_Sys[1].Cnv_Level[8].Cnv2.Inputs.VFD_Status := "C1208_StatusWord";
               "Control_DB".LCnv_Sys[1].Cnv_Level[8].Cnv2.Inputs.VFD_ActualCurrent := WORD_TO_INT("C1208_ActualCurrent");
               "Control_DB".LCnv_Sys[1].Cnv_Level[8].Cnv2.Inputs.VFD_Speed_Actual := WORD_TO_INT("C1208_ActualSpeed");
               "Control_DB".LCnv_Sys[1].Cnv_Level[8].Cnv2.Inputs.VFD_ActualTorque := "C1208_ActualTorque";
           END_REGION
       END_REGION

       REGION VTD
           "Control_DB".VTD_Sys[1].Inputs.Upper_Overtravel  := "OVERTRAVEL UPPER LIMIT - CH1(1)";
           "Control_DB".VTD_Sys[1].Inputs.Upper_limit := "VTD1 UPPER LIMIT";
           "Control_DB".VTD_Sys[1].Inputs.Ultimate_SlowDown := "VTD1 ULTIMATE SLOWDOWN";
           "Control_DB".VTD_Sys[1].Inputs.Ultimate_Creep := "VTD1 ULTIMATE CREEP";
           "Control_DB".VTD_Sys[1].Inputs.Lower_Limit := "VTD1 LOWER LIMIT";
           "Control_DB".VTD_Sys[1].Inputs.Lower_Overtravel := "OVERTRAVEL LOWER LIMIT - CH1(1)";
           "Control_DB".VTD_Sys[1].Inputs.Level_Detect1 := "VTD1 LEVEL DETECT 1";
           "Control_DB".VTD_Sys[1].Inputs.Level_Detect2 := "VTD1 LEVEL DETECT 2";
           "Control_DB".VTD_Sys[1].Inputs.DP1_Extended := "VTD1 DOCKING PINS EXTENDED 1";
           "Control_DB".VTD_Sys[1].Inputs.DP2_Extended := "VTD1 DOCKING PINS EXTENDED 2";
           "Control_DB".VTD_Sys[1].Inputs.DP1_Retracted := "VTD1 DOCKING PINS RETRACTED 1";
           "Control_DB".VTD_Sys[1].Inputs.DP2_Retracted := "VTD1 DOCKING PINS RETRACTED 2";
           "Control_DB".VTD_Sys[1].Inputs.Chain_Slack_1 := NOT "Remote_Panel_DB_1".Chain_Slack_1_Filtered;
           "Control_DB".VTD_Sys[1].Inputs.Chain_Slack_2 := NOT "Remote_Panel_DB_1".Chain_Slack_2_Filtered;
           "Control_DB".VTD_Sys[1].Inputs.Chain_Slack_3 := NOT "Remote_Panel_DB_1".Chain_Slack_3_Filtered;
           "Control_DB".VTD_Sys[1].Inputs.Chain_Slack_4 := NOT "Remote_Panel_DB_1".Chain_Slack_4_Filtered;
           "Control_DB".VTD_Sys[1].Inputs.PushToEnter := "VTD1 PUSH TO ENTER VTD ZONE";
           "Control_DB".VTD_Sys[1].Inputs.PushToExit := "VTD1 PUSH TO EXIT VTD ZONE";
           "Control_DB".VTD_Sys[1].Inputs.VFD_Status := "VTD1_StatusWord";
           "Control_DB".VTD_Sys[1].Inputs.VFD_ActualCurrent := REAL_TO_INT(("VTD1_ActualCurrent" / 10) / 72.5);
           "Control_DB".VTD_Sys[1].Inputs.VFD_Speed_Actual := "VTD1_ActualSpeed";
           "Control_DB".VTD_Sys[1].Inputs.VFD_ActualTorque := WORD_TO_INT("VTD1_ActualTorque");

       END_REGION

       REGION ABSOLUTE ENCODER
           REGION DOCUMENTATION
               //STATUS---------------------------------------------------------------------------------------------------------------------
               //
               //Encoder state word 2 - INPUT WORD 1
               //
               // 15 … 12 Encoder’s Sign-OF-Life (NOT relevant)
               // 11, 10 Reserved
               // 9 Control requested 0 = No control BY the PLC requested 1 = Control BY the PLC requested
               // 8 … 0 Reserved

               //Sensor 1 state word - INPUT WORD 2
               //
               // 15 Encoder error Description 0 = No error 1 = Error The error code is output in G1_XIST2.
               // 14 Park mode activated 0 = Normal operation 1 = Park mode activated Feedback based on G1_STW bit 14: No output OF position data G1_XIST1 AND G1_XIST2
               // 13 Transmission OF absolute position value 0 = No transmission 1 = Position value is output in G1_XIST2
               // 12 Status OF the Preset function (set/shift OF home position executed) 0 = No Preset function active 1 = Preset function is run Feedback based on G1_STW bit 12:  
               // 11 Requirement OF error acknowledgement detected New position value is output in G1_XIST1 AND G1_XIST2. On conclusion OF the Preset function the bit is set TO 0. 0 = No RETURN acknowledgement OF Encoder error 1 = Requirement OF error acknowledgement detected Reaction TO bit 15 in the sensor control word 1 G1_STW is acknowledged (see Table 14)
               // 10 Reserved
               // 9 … 0 NOT supported

               //Position 1 - INPUT WORD 3 AND 4
               // "AE_Position_1_Scaled" := (*SCALE_X(MIN := "Settings_DB".VTD_Settings.VTD_Min_Height,
               //                                   VALUE := *)NORM_X(MIN := 0,
               //                                                   VALUE := (SHL(IN:="AE_Position_1", N:=2) * 0.00228881) (*- "AE_Offset"*),
               //                                                   MAX := 1073741824)(*,
               //                                   MAX := "Settings_DB".VTD_Settings.VTD_Max_Heigh)*);
               // "mm_per_pulse" := 401,5584 / 262144;
               // 
               //CONTROL---------------------------------------------------------------------------------------------------------------------
               //
               //Encoder control word 2 - OUTPUT WORD 1
               //
               // 15 … 12 Master’s Sign-OF-Life (NOT relevant)
               // 10 control BY PLC 0 = No control BY the PLC 1 = Control BY the PLC Enables the PLC BY using control words TO activate / deactivate encoder functions
               // 7 Fault acknowledge Error-buffer handling NOT supported
               // 11, 9, 8, 6 … 0 Reserved
               // "AE_Control_Word_1".%X10 := "AE_PLC_Control";
               // 
               //Sensor 1 control word - OUTPUT WORD 2-------------------------------------------------------------------------------------------
               //
               // 15 Acknowledging a sensor error Description 0 = Encoder error message NOT acknowledged BY PLC 1 = Encoder error message acknowledged BY the PLC
               // 14 Activate park mode 0 = Normal operation 1 = Activate park mode
               // 13 Request FOR the absolute position value 0 = No request 1 = Request BY the master Results in the cyclic output OF the position values in G1_XIST2
               // 12 Activate preset value (see note below) Defines that a configured preset value is used (see section 3.5 on page 24) 0 = Preset value is NOT activated 1 = Preset value is activated
               // 11 Preset mode Defines how a configured preset value is used 0 = Preset value is used as a new absolute value 1 = Preset value is added TO the previous value
               // 10 … 0 Reserved
               // "AE_Control_Word_2".%X15 := "VTD_Reset_HMI_Tags";
               // "AE_Control_Word_2".%X14 := "AE_Activate_ParkMode";
               // "AE_Control_Word_2".%X13 := "AE_Request_ABS_Value";
               // "AE_Control_Word_2".%X12 := "AE_Activate_Preset_Value";
               // "AE_Control_Word_2".%X11 := "AE_Preset_Mode";
           END_REGION

           //STATUS---------------------------------------------------------------------------------------------------------------------
           "Control_DB".VTD_Sys[1].Inputs.AE_Status_2 := "AE_Status_2(1)";
           //Position 1 - INPUT WORD 3 AND 4
           "Control_DB".VTD_Sys[1].Inputs.AE_Position_1 := REAL_TO_DINT(((((*1073741823 - reverse the direction*)
    (SHR(IN := "AE_Position_1(1)", N := 2))) - 31381317) * 0.0015318237304688 (*Mechanical relationship*)+ 48062)(*Offset*));

           // Position 2 - INPUT WORD 5 AND 6
           "Control_DB".VTD_Sys[1].Inputs.AE_Position_2 := SHR(IN := "AE_Position_2(1)", N := 2);

           //Speed A - INPUT WORD 7
           "Control_DB".VTD_Sys[1].Inputs.AE_Speed := "AE_Speed(1)" * 10;
       END_REGION

       REGION LINEAR ENCODER
           "Control_DB".VTD_Sys[1].Inputs.LE_Position := "LE_X_Unsafe_Position(1)" / 10;
           "Control_DB".VTD_Sys[1].Inputs.LE_Speed := "LE_Speed(1)" * 100;
           "Control_DB".VTD_Sys[1].Inputs.LE_Status := "LE_Status(1)";
           "Control_DB".VTD_Sys[1].Inputs.LE_Warnings := "LE_Warnings(1)";
           REGION DOCUMENTATION
               //STATUS 
               //
               // 0 ERR - Error message (Error code in XP00– XP15); remaining bits = 0, see Error Codes
               // 1 NP - No position information/OUT (XP = 0, YP = 0, SP = 0)
               // 2 WRN - Warnings present, see Warning Module
               // 3 EV - Event present
               // 4 posdetected - Valid position information available

               //WARNINGS
               //
               // 0 WRN01 A code with non-PXV content was found.
               // 1 WRN02 the read head is too close TO the Data Matrix code tape.
               // 2 WRN03 the read head is too far from the Data Matrix code tape.
               // 3 WRN04 Y position too large. The sensor is just before OUT.
               // 4 WRN05 Y position is too small. The sensor is just before OUT.
               // 5 WRN06 the read head is rotated OR tilted in relation TO the Data Matrix code tape.
               // 6 WRN07 Low level OF code contrast.
               // 7 WRN08 Repair tape detected.
               // 8 WRN09 Temperature too high.
               // 9...15 Reserved

               //QUALITY GRADE
               //
               //The quality grades enable constant monitoring of the code tape and the camera along the entire
               //traverse distance. This enables you to detect and act upon potential damage or contamination
               //of the code tape and camera at the earliest stage possible during commissioning and normal
               //operation. As a result, this maximizes the overall functional reliability of your plant, and
               //it means you are able to immediately localize the issue in the case of a fault. Evaluations
               //are made using a scale of 1 to 6. The value 1 is the best possible read quality. A value greater
               //than 3 or worse requires the camera and its path to be inspected. The value 7 signifies "No position"
               //because no code was detected. An evaluation that indicates poor quality as the outcome can be due to
               //a misalignment or incorrect orientation, an incorrect measuring distance, or because the code tape has been affixed incorrectly
           END_REGION
       END_REGION

       REGION SICK BARCODE LECTORS
           IF "Control_DB".VTDBarcode_Station[1].Running AND "SICK_Lector_Control_DB_1".Result <> "Control_DB".VTDBarcode_Station[1].Barcode_Old THEN
               "Control_DB".VTD_Sys[1].Inputs."Barcode 1" := "SICK_Lector_Control_DB_1".Result;
               // "Control_DB".VTD_Control.Inputs."Barcode 2'" := SICK_Barcode_DB".Result;
               // "Control_DB".VTDBarcode_Station[1].Barcode_Old := "SICK_Lector_DB_1".Barcode_Result;
           ELSE
               "Control_DB".VTD_Sys[1].Inputs."Barcode 1" :=
               "Control_DB".VTD_Sys[1].Inputs."Barcode 2" := '';
           END_IF;

       END_REGION

       REGION VFD HARDWARE ID
           //Buffer conveyors 1
           "Settings_DB".LCnv_Sys[1].Cnv_Level[1].Cnv1.G120_Hardware_ID := "C1101~Drive_1~Standard_telegram_20__PZD-2_6";
           "Settings_DB".LCnv_Sys[1].Cnv_Level[2].Cnv1.G120_Hardware_ID := "C1102~Drive_1~Standard_telegram_20__PZD-2_6";
           "Settings_DB".LCnv_Sys[1].Cnv_Level[3].Cnv1.G120_Hardware_ID := "C1103~Drive_1~Standard_telegram_20__PZD-2_6";
           "Settings_DB".LCnv_Sys[1].Cnv_Level[4].Cnv1.G120_Hardware_ID := "C1104~Drive_1~Standard_telegram_20__PZD-2_6";
           "Settings_DB".LCnv_Sys[1].Cnv_Level[5].Cnv1.G120_Hardware_ID := "C1105~Drive_1~Standard_telegram_20__PZD-2_6";
           "Settings_DB".LCnv_Sys[1].Cnv_Level[6].Cnv1.G120_Hardware_ID := "C1106~Drive_1~Standard_telegram_20__PZD-2_6";
           "Settings_DB".LCnv_Sys[1].Cnv_Level[7].Cnv1.G120_Hardware_ID := "C1107~Drive_1~Standard_telegram_20__PZD-2_6";
           "Settings_DB".LCnv_Sys[1].Cnv_Level[8].Cnv1.G120_Hardware_ID := "C1108~Drive_1~Standard_telegram_20__PZD-2_6";

           //Buffer conveyors 2
           "Settings_DB".LCnv_Sys[1].Cnv_Level[1].Cnv2.G120_Hardware_ID := "C1201~Drive_1~Standard_telegram_20__PZD-2_6";
           "Settings_DB".LCnv_Sys[1].Cnv_Level[2].Cnv2.G120_Hardware_ID := "C1202~Drive_1~Standard_telegram_20__PZD-2_6";
           "Settings_DB".LCnv_Sys[1].Cnv_Level[3].Cnv2.G120_Hardware_ID := "C1203~Drive_1~Standard_telegram_20__PZD-2_6";
           "Settings_DB".LCnv_Sys[1].Cnv_Level[4].Cnv2.G120_Hardware_ID := "C1204~Drive_1~Standard_telegram_20__PZD-2_6";
           "Settings_DB".LCnv_Sys[1].Cnv_Level[5].Cnv2.G120_Hardware_ID := "C1205~Drive_1~Standard_telegram_20__PZD-2_6";
           "Settings_DB".LCnv_Sys[1].Cnv_Level[6].Cnv2.G120_Hardware_ID := "C1206~Drive_1~Standard_telegram_20__PZD-2_6";
           "Settings_DB".LCnv_Sys[1].Cnv_Level[7].Cnv2.G120_Hardware_ID := "C1207~Drive_1~Standard_telegram_20__PZD-2_6";
           "Settings_DB".LCnv_Sys[1].Cnv_Level[8].Cnv2.G120_Hardware_ID := "C1208~Drive_1~Standard_telegram_20__PZD-2_6";

           //Extractor conveyor
           "Settings_DB".ECnv_Sys[1].G120_Hardware_ID := "CVTD_1~Drive_1~Standard_telegram_20__PZD-2_6";

           //VTD
           "Settings_DB".VTD_Sys[1].G120_Hardware_ID := "VTD_1~DO_VECTOR_1~Standard_telegram_20__PZD-2_6";
       END_REGION
   END_REGION

   REGION SYSTEM 2
       REGION EXTRACTOR CONVEYOR
           "Control_DB".ECnv_Sys[2].Inputs.Left := "CVTD2 SENSOR CONVEYOR LEFT";
           "Control_DB".ECnv_Sys[2].Inputs.Lpd1 := "CVTD2 SENSOR CONVEYOR LEFT (PALLET DETECT 1)";
           "Control_DB".ECnv_Sys[2].Inputs.Center := "CVTD2 SENSOR CONVEYOR CENTER";
           "Control_DB".ECnv_Sys[2].Inputs.Right := "CVTD2 SENSOR CONVEYOR RIGHT";
           "Control_DB".ECnv_Sys[2].Inputs.Rpd1 := "CVTD2 SENSOR CONVEYOR RIGHT (PALLET DETECT 1)";

           "T_OH_Left_2".TOF(IN := "CVTD2 OVERHANG LEFT" OR NOT "Control_DB".VTD_Sys[2].Running,
                             PT := T#200ms);
           "Control_DB".ECnv_Sys[2].Inputs.Overhang_Left := "T_OH_Left_2".Q;

           "T_OH_Right_2".TOF(IN:= "CVTD2 OVERHANG RIGHT" OR NOT "Control_DB".VTD_Sys[2].Running,
                             PT:= T#200ms);
          "Control_DB".ECnv_Sys[2].Inputs.Overhang_Right := "T_OH_Right_2".Q;

           "Control_DB".ECnv_Sys[2].Inputs.VFD_Status := "CVTD2_StatusWord";
           "Control_DB".ECnv_Sys[2].Inputs.VFD_ActualCurrent := WORD_TO_INT("CVTD2_ActualCurrent");
           "Control_DB".ECnv_Sys[2].Inputs.VFD_Speed_Actual := WORD_TO_INT("CVTD2_ActualSpeed");
           "Control_DB".ECnv_Sys[2].Inputs.VFD_ActualTorque := WORD_TO_INT("CVTD2_ActualTorque");
       END_REGION

       REGION BUFFER CONVEYORS
           REGION LEVEL 1
               //BUFFER CONVEYOR LEVEL 1 - CONVEYOR 1
               "Control_DB".LCnv_Sys[2].Cnv_Level[1].Cnv1.Inputs.Left := NOT "C2101 - SENSOR CNV LEFT";
               "Control_DB".LCnv_Sys[2].Cnv_Level[1].Cnv1.Inputs.Lpd1 := NOT "C2101 - SENSOR CNV LEFT (PALLET DETECT 1)";
               "Control_DB".LCnv_Sys[2].Cnv_Level[1].Cnv1.Inputs.Lpd2 := NOT "C2101 - SENSOR CNV LEFT (PALLET DETECT 2)";
               "Control_DB".LCnv_Sys[2].Cnv_Level[1].Cnv1.Inputs.Right := NOT "C2101 - SENSOR CNV RIGHT";
               "Control_DB".LCnv_Sys[2].Cnv_Level[1].Cnv1.Inputs.Rpd1 := NOT "C2101 - SENSOR CNV RIGHT (PALLET DETECT 1)";
               "Control_DB".LCnv_Sys[2].Cnv_Level[1].Cnv1.Inputs.Rpd2 := NOT "C2101 - SENSOR CNV RIGHT (PALLET DETECT 2)";
               "Control_DB".LCnv_Sys[2].Cnv_Level[1].Cnv1.Inputs.Sdetect1 := NOT "C2101 - SHUTTLE IN POSITION 1";
               "Control_DB".LCnv_Sys[2].Cnv_Level[1].Cnv1.Inputs.Sdetect2 := NOT "C2101 - SHUTTLE IN POSITION 2";

               "Control_DB".LCnv_Sys[2].Cnv_Level[1].Cnv1.Inputs.VFD_Status := "C2101_StatusWord";
               "Control_DB".LCnv_Sys[2].Cnv_Level[1].Cnv1.Inputs.VFD_ActualCurrent :=WORD_TO_INT("C2101_ActualCurrent");
               "Control_DB".LCnv_Sys[2].Cnv_Level[1].Cnv1.Inputs.VFD_Speed_Actual :=WORD_TO_INT("C2101_ActualSpeed");
               "Control_DB".LCnv_Sys[2].Cnv_Level[1].Cnv1.Inputs.VFD_ActualTorque := WORD_TO_INT("C2101_ActualTorque");

               //BUFFER CONVEYOR LEVEL 1 - CONVEYOR 2
               "Control_DB".LCnv_Sys[2].Cnv_Level[1].Cnv2.Inputs.Left := NOT "C2201 - SENSOR CNV LEFT";
               "Control_DB".LCnv_Sys[2].Cnv_Level[1].Cnv2.Inputs.Lpd1 := NOT "C2201 - SENSOR CNV LEFT (PALLET DETECT 1)";
               "Control_DB".LCnv_Sys[2].Cnv_Level[1].Cnv2.Inputs.Lpd2 := NOT "C2201 - SENSOR CNV LEFT (PALLET DETECT 2)";
               "Control_DB".LCnv_Sys[2].Cnv_Level[1].Cnv2.Inputs.Right := NOT "C2201 - SENSOR CNV RIGHT";
               "Control_DB".LCnv_Sys[2].Cnv_Level[1].Cnv2.Inputs.Rpd1 := NOT "C2201 - SENSOR CNV RIGHT (PALLET DETECT 1)";
               "Control_DB".LCnv_Sys[2].Cnv_Level[1].Cnv2.Inputs.Rpd2 := NOT "C2201 - SENSOR CNV RIGHT (PALLET DETECT 2)";
               "Control_DB".LCnv_Sys[2].Cnv_Level[1].Cnv2.Inputs.Sdetect1 := NOT "C2201 - SHUTTLE IN POSITION 1";
               "Control_DB".LCnv_Sys[2].Cnv_Level[1].Cnv2.Inputs.Sdetect2 := NOT "C2201 - SHUTTLE IN POSITION 2";

               "Control_DB".LCnv_Sys[2].Cnv_Level[1].Cnv2.Inputs.VFD_Status := "C2201_StatusWord";
               "Control_DB".LCnv_Sys[2].Cnv_Level[1].Cnv2.Inputs.VFD_ActualCurrent := WORD_TO_INT("C2201_ActualCurrent");
               "Control_DB".LCnv_Sys[2].Cnv_Level[1].Cnv2.Inputs.VFD_Speed_Actual := WORD_TO_INT("C2201_ActualSpeed");
               "Control_DB".LCnv_Sys[2].Cnv_Level[1].Cnv2.Inputs.VFD_ActualTorque := WORD_TO_INT("C2201_ActualTorque");
           END_REGION

           REGION LEVEL 2
               //BUFFER CONVEYOR LEVEL 2 - CONVEYOR 1
               "Control_DB".LCnv_Sys[2].Cnv_Level[2].Cnv1.Inputs.Left := NOT "C2102 - SENSOR CNV LEFT";
               "Control_DB".LCnv_Sys[2].Cnv_Level[2].Cnv1.Inputs.Lpd1 := NOT "C2102 - SENSOR CNV LEFT (PALLET DETECT 1)";
               "Control_DB".LCnv_Sys[2].Cnv_Level[2].Cnv1.Inputs.Lpd2 := NOT "C2102 - SENSOR CNV LEFT (PALLET DETECT 2)";
               "Control_DB".LCnv_Sys[2].Cnv_Level[2].Cnv1.Inputs.Right := NOT "C2102 - SENSOR CNV RIGHT";
               "Control_DB".LCnv_Sys[2].Cnv_Level[2].Cnv1.Inputs.Rpd1 := NOT "C2102 - SENSOR CNV RIGHT (PALLET DETECT 1)";
               "Control_DB".LCnv_Sys[2].Cnv_Level[2].Cnv1.Inputs.Rpd2 := NOT "C2102 - SENSOR CNV RIGHT (PALLET DETECT 2)";
               "Control_DB".LCnv_Sys[2].Cnv_Level[2].Cnv1.Inputs.Sdetect1 := NOT "C2102 - SHUTTLE IN POSITION 1";
               "Control_DB".LCnv_Sys[2].Cnv_Level[2].Cnv1.Inputs.Sdetect2 := NOT "C2102 - SHUTTLE IN POSITION 2";
               "Control_DB".LCnv_Sys[2].Cnv_Level[2].Cnv1.Safety_Stop_Cnrl.Inputs.DP_Extended := "C2102 - SENSOR SAFETY PIN1 UP";
               "Control_DB".LCnv_Sys[2].Cnv_Level[2].Cnv1.Safety_Stop_Cnrl.Inputs.DP_Retracted := "C2102 - SENSOR SAFETY PIN1 DOWN";

               "Control_DB".LCnv_Sys[2].Cnv_Level[2].Cnv1.Inputs.VFD_Status := "C2102_StatusWord";
               "Control_DB".LCnv_Sys[2].Cnv_Level[2].Cnv1.Inputs.VFD_ActualCurrent := WORD_TO_INT("C2102_ActualCurrent");
               "Control_DB".LCnv_Sys[2].Cnv_Level[2].Cnv1.Inputs.VFD_Speed_Actual := WORD_TO_INT("C2102_ActualSpeed");
               "Control_DB".LCnv_Sys[2].Cnv_Level[2].Cnv1.Inputs.VFD_ActualTorque := WORD_TO_INT("C2102_ActualTorque");

               //BUFFER CONVEYOR LEVEL 2 - CONVEYOR 2
               "Control_DB".LCnv_Sys[2].Cnv_Level[2].Cnv2.Inputs.Left := NOT "C2202 - SENSOR CNV LEFT";
               "Control_DB".LCnv_Sys[2].Cnv_Level[2].Cnv2.Inputs.Lpd1 := NOT "C2202 - SENSOR CNV LEFT (PALLET DETECT 1)";
               "Control_DB".LCnv_Sys[2].Cnv_Level[2].Cnv2.Inputs.Lpd2 := NOT "C2202 - SENSOR CNV LEFT (PALLET DETECT 2)";
               "Control_DB".LCnv_Sys[2].Cnv_Level[2].Cnv2.Inputs.Right := NOT "C2202 - SENSOR CNV RIGHT";
               "Control_DB".LCnv_Sys[2].Cnv_Level[2].Cnv2.Inputs.Rpd1 := NOT "C2202 - SENSOR CNV RIGHT (PALLET DETECT 1)";
               "Control_DB".LCnv_Sys[2].Cnv_Level[2].Cnv2.Inputs.Rpd2 := NOT "C2202 - SENSOR CNV RIGHT (PALLET DETECT 2)";
               "Control_DB".LCnv_Sys[2].Cnv_Level[2].Cnv2.Inputs.Sdetect1 := NOT "C2202 - SHUTTLE IN POSITION 1";
               "Control_DB".LCnv_Sys[2].Cnv_Level[2].Cnv2.Inputs.Sdetect2 := NOT "C2202 - SHUTTLE IN POSITION 2";
               "Control_DB".LCnv_Sys[2].Cnv_Level[2].Cnv2.Safety_Stop_Cnrl.Inputs.DP_Extended := "C2202 - SENSOR SAFETY PIN1 UP";
               "Control_DB".LCnv_Sys[2].Cnv_Level[2].Cnv2.Safety_Stop_Cnrl.Inputs.DP_Retracted := "C2202 - SENSOR SAFETY PIN1 DOWN";

               "Control_DB".LCnv_Sys[2].Cnv_Level[2].Cnv2.Inputs.VFD_Status := "C2202_StatusWord";
               "Control_DB".LCnv_Sys[2].Cnv_Level[2].Cnv2.Inputs.VFD_ActualCurrent := WORD_TO_INT("C2202_ActualCurrent");
               "Control_DB".LCnv_Sys[2].Cnv_Level[2].Cnv2.Inputs.VFD_Speed_Actual := WORD_TO_INT("C2202_ActualSpeed");
               "Control_DB".LCnv_Sys[2].Cnv_Level[2].Cnv2.Inputs.VFD_ActualTorque := WORD_TO_INT("C2202_ActualTorque");
           END_REGION

           REGION LEVEL 3
               //BUFFER CONVEYOR LEVEL 3 - CONVEYOR 1
               "Control_DB".LCnv_Sys[2].Cnv_Level[3].Cnv1.Inputs.Left := NOT "C2103 - SENSOR CNV LEFT";
               "Control_DB".LCnv_Sys[2].Cnv_Level[3].Cnv1.Inputs.Lpd1 := NOT "C2103 - SENSOR CNV LEFT (PALLET DETECT 1)";
               "Control_DB".LCnv_Sys[2].Cnv_Level[3].Cnv1.Inputs.Lpd2 := NOT "C2103 - SENSOR CNV LEFT (PALLET DETECT 2)";
               "Control_DB".LCnv_Sys[2].Cnv_Level[3].Cnv1.Inputs.Right := NOT "C2103 - SENSOR CNV RIGHT";
               "Control_DB".LCnv_Sys[2].Cnv_Level[3].Cnv1.Inputs.Rpd1 := NOT "C2103 - SENSOR CNV RIGHT (PALLET DETECT 1)";
               "Control_DB".LCnv_Sys[2].Cnv_Level[3].Cnv1.Inputs.Rpd2 := NOT "C2103 - SENSOR CNV RIGHT (PALLET DETECT 2)";
               "Control_DB".LCnv_Sys[2].Cnv_Level[3].Cnv1.Inputs.Sdetect1 := NOT "C2103 - SHUTTLE IN POSITION 1";
               "Control_DB".LCnv_Sys[2].Cnv_Level[3].Cnv1.Inputs.Sdetect2 := NOT "C2103 - SHUTTLE IN POSITION 2";
               "Control_DB".LCnv_Sys[2].Cnv_Level[3].Cnv1.Safety_Stop_Cnrl.Inputs.DP_Extended := "C2103 - SENSOR SAFETY PIN1 UP";
               "Control_DB".LCnv_Sys[2].Cnv_Level[3].Cnv1.Safety_Stop_Cnrl.Inputs.DP_Retracted := "C2103 - SENSOR SAFETY PIN1 DOWN";

               "Control_DB".LCnv_Sys[2].Cnv_Level[3].Cnv1.Inputs.VFD_Status := "C2103_StatusWord";
               "Control_DB".LCnv_Sys[2].Cnv_Level[3].Cnv1.Inputs.VFD_ActualCurrent := WORD_TO_INT("C2103_ActualCurrent");
               "Control_DB".LCnv_Sys[2].Cnv_Level[3].Cnv1.Inputs.VFD_Speed_Actual := WORD_TO_INT("C2103_ActualSpeed");
               "Control_DB".LCnv_Sys[2].Cnv_Level[3].Cnv1.Inputs.VFD_ActualTorque := WORD_TO_INT("C2103_ActualTorque");

               //BUFFER CONVEYOR LEVEL 3 - CONVEYOR 2
               "Control_DB".LCnv_Sys[2].Cnv_Level[3].Cnv2.Inputs.Left := NOT "C2203 - SENSOR CNV LEFT";
               "Control_DB".LCnv_Sys[2].Cnv_Level[3].Cnv2.Inputs.Lpd1 := NOT "C2203 - SENSOR CNV LEFT (PALLET DETECT 1)";
               "Control_DB".LCnv_Sys[2].Cnv_Level[3].Cnv2.Inputs.Lpd2 := NOT "C2203 - SENSOR CNV LEFT (PALLET DETECT 2)";
               "Control_DB".LCnv_Sys[2].Cnv_Level[3].Cnv2.Inputs.Right := NOT "C2203 - SENSOR CNV RIGHT";
               "Control_DB".LCnv_Sys[2].Cnv_Level[3].Cnv2.Inputs.Rpd1 := NOT "C2203 - SENSOR CNV RIGHT (PALLET DETECT 1)";
               "Control_DB".LCnv_Sys[2].Cnv_Level[3].Cnv2.Inputs.Rpd2 := NOT "C2203 - SENSOR CNV RIGHT (PALLET DETECT 2)";
               "Control_DB".LCnv_Sys[2].Cnv_Level[3].Cnv2.Inputs.Sdetect1 := NOT "C2203 - SHUTTLE IN POSITION 1";
               "Control_DB".LCnv_Sys[2].Cnv_Level[3].Cnv2.Inputs.Sdetect2 := NOT "C2203 - SHUTTLE IN POSITION 2";
               "Control_DB".LCnv_Sys[2].Cnv_Level[3].Cnv2.Safety_Stop_Cnrl.Inputs.DP_Extended := "C2203 - SENSOR SAFETY PIN1 UP";
               "Control_DB".LCnv_Sys[2].Cnv_Level[3].Cnv2.Safety_Stop_Cnrl.Inputs.DP_Retracted := "C2203 - SENSOR SAFETY PIN1 DOWN";

               "Control_DB".LCnv_Sys[2].Cnv_Level[3].Cnv2.Inputs.VFD_Status := "C2203_StatusWord";
               "Control_DB".LCnv_Sys[2].Cnv_Level[3].Cnv2.Inputs.VFD_ActualCurrent := WORD_TO_INT("C2203_ActualCurrent");
               "Control_DB".LCnv_Sys[2].Cnv_Level[3].Cnv2.Inputs.VFD_Speed_Actual := WORD_TO_INT("C2203_ActualSpeed");
           END_REGION

           REGION LEVEL 4
               //BUFFER CONVEYOR LEVEL 4 - CONVEYOR 1
               "Control_DB".LCnv_Sys[2].Cnv_Level[4].Cnv1.Inputs.Left := NOT "C2104 - SENSOR CNV LEFT";
               "Control_DB".LCnv_Sys[2].Cnv_Level[4].Cnv1.Inputs.Lpd1 := NOT "C2104 - SENSOR CNV LEFT (PALLET DETECT 1)";
               "Control_DB".LCnv_Sys[2].Cnv_Level[4].Cnv1.Inputs.Lpd2 := NOT "C2104 - SENSOR CNV LEFT (PALLET DETECT 2)";
               "Control_DB".LCnv_Sys[2].Cnv_Level[4].Cnv1.Inputs.Right := NOT "C2104 - SENSOR CNV RIGHT";
               "Control_DB".LCnv_Sys[2].Cnv_Level[4].Cnv1.Inputs.Rpd1 := NOT "C2104 - SENSOR CNV RIGHT (PALLET DETECT 1)";
               "Control_DB".LCnv_Sys[2].Cnv_Level[4].Cnv1.Inputs.Rpd2 := NOT "C2104 - SENSOR CNV RIGHT (PALLET DETECT 2)";
               "Control_DB".LCnv_Sys[2].Cnv_Level[4].Cnv1.Inputs.Sdetect1 := NOT "C2104 - SHUTTLE IN POSITION 1";
               "Control_DB".LCnv_Sys[2].Cnv_Level[4].Cnv1.Inputs.Sdetect2 := NOT "C2104 - SHUTTLE IN POSITION 2";
               "Control_DB".LCnv_Sys[2].Cnv_Level[4].Cnv1.Safety_Stop_Cnrl.Inputs.DP_Extended := "C2104 - SENSOR SAFETY PIN1 UP";
               "Control_DB".LCnv_Sys[2].Cnv_Level[4].Cnv1.Safety_Stop_Cnrl.Inputs.DP_Retracted := "C2104 - SENSOR SAFETY PIN1 DOWN";

               "Control_DB".LCnv_Sys[2].Cnv_Level[4].Cnv1.Inputs.VFD_Status := "C2104_StatusWord";
               "Control_DB".LCnv_Sys[2].Cnv_Level[4].Cnv1.Inputs.VFD_ActualCurrent := WORD_TO_INT("C2104_ActualCurrent");
               "Control_DB".LCnv_Sys[2].Cnv_Level[4].Cnv1.Inputs.VFD_Speed_Actual := WORD_TO_INT("C2104_ActualSpeed");
               "Control_DB".LCnv_Sys[2].Cnv_Level[4].Cnv1.Inputs.VFD_ActualTorque := WORD_TO_INT("C2104_ActualTorque");

               //BUFFER CONVEYOR LEVEL 4 - CONVEYOR 2
               "Control_DB".LCnv_Sys[2].Cnv_Level[4].Cnv2.Inputs.Left := NOT "C2204 - SENSOR CNV LEFT";
               "Control_DB".LCnv_Sys[2].Cnv_Level[4].Cnv2.Inputs.Lpd1 := NOT "C2204 - SENSOR CNV LEFT (PALLET DETECT 1)";
               "Control_DB".LCnv_Sys[2].Cnv_Level[4].Cnv2.Inputs.Lpd2 := NOT "C2204 - SENSOR CNV LEFT (PALLET DETECT 2)";
               "Control_DB".LCnv_Sys[2].Cnv_Level[4].Cnv2.Inputs.Right := NOT "C2204 - SENSOR CNV RIGHT";
               "Control_DB".LCnv_Sys[2].Cnv_Level[4].Cnv2.Inputs.Rpd1 := NOT "C2204 - SENSOR CNV RIGHT (PALLET DETECT 1)";
               "Control_DB".LCnv_Sys[2].Cnv_Level[4].Cnv2.Inputs.Rpd2 := NOT "C2204 - SENSOR CNV RIGHT (PALLET DETECT 2)";
               "Control_DB".LCnv_Sys[2].Cnv_Level[4].Cnv2.Inputs.Sdetect1 := NOT "C2204 - SHUTTLE IN POSITION 1";
               "Control_DB".LCnv_Sys[2].Cnv_Level[4].Cnv2.Inputs.Sdetect2 := NOT "C2204 - SHUTTLE IN POSITION 2";
               "Control_DB".LCnv_Sys[2].Cnv_Level[4].Cnv2.Safety_Stop_Cnrl.Inputs.DP_Extended := "C2204 - SENSOR SAFETY PIN1 UP";
               "Control_DB".LCnv_Sys[2].Cnv_Level[4].Cnv2.Safety_Stop_Cnrl.Inputs.DP_Retracted := "C2204 - SENSOR SAFETY PIN1 DOWN";

               "Control_DB".LCnv_Sys[2].Cnv_Level[4].Cnv2.Inputs.VFD_Status := "C2204_StatusWord";
               "Control_DB".LCnv_Sys[2].Cnv_Level[4].Cnv2.Inputs.VFD_ActualCurrent := WORD_TO_INT("C2204_ActualCurrent");
               "Control_DB".LCnv_Sys[2].Cnv_Level[4].Cnv2.Inputs.VFD_Speed_Actual := WORD_TO_INT("C2204_ActualSpeed");
               "Control_DB".LCnv_Sys[2].Cnv_Level[4].Cnv2.Inputs.VFD_ActualTorque := WORD_TO_INT("C2204_ActualTorque");
           END_REGION

           REGION LEVEL 5
               //BUFFER CONVEYOR LEVEL 5 - CONVEYOR 1
               "Control_DB".LCnv_Sys[2].Cnv_Level[5].Cnv1.Inputs.Left := NOT "C2105 - SENSOR CNV LEFT";
               "Control_DB".LCnv_Sys[2].Cnv_Level[5].Cnv1.Inputs.Lpd1 := NOT "C2105 - SENSOR CNV LEFT (PALLET DETECT 1)";
               "Control_DB".LCnv_Sys[2].Cnv_Level[5].Cnv1.Inputs.Lpd2 := NOT "C2105 - SENSOR CNV LEFT (PALLET DETECT 2)";
               "Control_DB".LCnv_Sys[2].Cnv_Level[5].Cnv1.Inputs.Right := NOT "C2105 - SENSOR CNV RIGHT";
               "Control_DB".LCnv_Sys[2].Cnv_Level[5].Cnv1.Inputs.Rpd1 := NOT "C2105 - SENSOR CNV RIGHT (PALLET DETECT 1)";
               "Control_DB".LCnv_Sys[2].Cnv_Level[5].Cnv1.Inputs.Rpd2 := NOT "C2105 - SENSOR CNV RIGHT (PALLET DETECT 2)";
               "Control_DB".LCnv_Sys[2].Cnv_Level[5].Cnv1.Inputs.Sdetect1 := NOT "C2105 - SHUTTLE IN POSITION 1";
               "Control_DB".LCnv_Sys[2].Cnv_Level[5].Cnv1.Inputs.Sdetect2 := NOT "C2105 - SHUTTLE IN POSITION 2";
               "Control_DB".LCnv_Sys[2].Cnv_Level[5].Cnv1.Safety_Stop_Cnrl.Inputs.DP_Extended := "C2105 - SENSOR SAFETY PIN1 UP";
               "Control_DB".LCnv_Sys[2].Cnv_Level[5].Cnv1.Safety_Stop_Cnrl.Inputs.DP_Retracted := "C2105 - SENSOR SAFETY PIN1 DOWN";

               "Control_DB".LCnv_Sys[2].Cnv_Level[5].Cnv1.Inputs.VFD_Status := "C2105_StatusWord";
               "Control_DB".LCnv_Sys[2].Cnv_Level[5].Cnv1.Inputs.VFD_ActualCurrent := WORD_TO_INT("C2105_ActualCurrent");
               "Control_DB".LCnv_Sys[2].Cnv_Level[5].Cnv1.Inputs.VFD_Speed_Actual := WORD_TO_INT("C2105_ActualSpeed");
               "Control_DB".LCnv_Sys[2].Cnv_Level[5].Cnv1.Inputs.VFD_ActualTorque := WORD_TO_INT("C2105_ActualTorque");

               //BUFFER CONVEYOR LEVEL 5 - CONVEYOR 2
               "Control_DB".LCnv_Sys[2].Cnv_Level[5].Cnv2.Inputs.Left := NOT "C2205 - SENSOR CNV LEFT";
               "Control_DB".LCnv_Sys[2].Cnv_Level[5].Cnv2.Inputs.Lpd1 := NOT "C2205 - SENSOR CNV LEFT (PALLET DETECT 1)";
               "Control_DB".LCnv_Sys[2].Cnv_Level[5].Cnv2.Inputs.Lpd2 := NOT "C2205 - SENSOR CNV LEFT (PALLET DETECT 2)";
               "Control_DB".LCnv_Sys[2].Cnv_Level[5].Cnv2.Inputs.Right := NOT "C2205 - SENSOR CNV RIGHT";
               "Control_DB".LCnv_Sys[2].Cnv_Level[5].Cnv2.Inputs.Rpd1 := NOT "C2205 - SENSOR CNV RIGHT (PALLET DETECT 1)";
               "Control_DB".LCnv_Sys[2].Cnv_Level[5].Cnv2.Inputs.Rpd2 := NOT "C2205 - SENSOR CNV RIGHT (PALLET DETECT 2)";
               "Control_DB".LCnv_Sys[2].Cnv_Level[5].Cnv2.Inputs.Sdetect1 := NOT "C2205 - SHUTTLE IN POSITION 1";
               "Control_DB".LCnv_Sys[2].Cnv_Level[5].Cnv2.Inputs.Sdetect2 := NOT "C2205 - SHUTTLE IN POSITION 2";
               "Control_DB".LCnv_Sys[2].Cnv_Level[5].Cnv2.Safety_Stop_Cnrl.Inputs.DP_Extended := "C2205 - SENSOR SAFETY PIN1 UP";
               "Control_DB".LCnv_Sys[2].Cnv_Level[5].Cnv2.Safety_Stop_Cnrl.Inputs.DP_Retracted := "C2205 - SENSOR SAFETY PIN1 DOWN";

               "Control_DB".LCnv_Sys[2].Cnv_Level[5].Cnv2.Inputs.VFD_Status := "C2205_StatusWord";
               "Control_DB".LCnv_Sys[2].Cnv_Level[5].Cnv2.Inputs.VFD_ActualCurrent := WORD_TO_INT("C2205_ActualCurrent");
               "Control_DB".LCnv_Sys[2].Cnv_Level[5].Cnv2.Inputs.VFD_Speed_Actual := WORD_TO_INT("C2205_ActualSpeed");
               "Control_DB".LCnv_Sys[2].Cnv_Level[5].Cnv2.Inputs.VFD_ActualTorque := WORD_TO_INT("C2205_ActualTorque");
           END_REGION

           REGION LEVEL 6
               //BUFFER CONVEYOR LEVEL 6 - CONVEYOR 1
               "Control_DB".LCnv_Sys[2].Cnv_Level[6].Cnv1.Inputs.Left := NOT "C2106 - SENSOR CNV LEFT";
               "Control_DB".LCnv_Sys[2].Cnv_Level[6].Cnv1.Inputs.Lpd1 := NOT "C2106 - SENSOR CNV LEFT (PALLET DETECT 1)";
               "Control_DB".LCnv_Sys[2].Cnv_Level[6].Cnv1.Inputs.Lpd2 := NOT "C2106 - SENSOR CNV LEFT (PALLET DETECT 2)";
               "Control_DB".LCnv_Sys[2].Cnv_Level[6].Cnv1.Inputs.Right := NOT "C2106 - SENSOR CNV RIGHT";
               "Control_DB".LCnv_Sys[2].Cnv_Level[6].Cnv1.Inputs.Rpd1 := NOT "C2106 - SENSOR CNV RIGHT (PALLET DETECT 1)";
               "Control_DB".LCnv_Sys[2].Cnv_Level[6].Cnv1.Inputs.Rpd2 := NOT "C2106 - SENSOR CNV RIGHT (PALLET DETECT 2)";
               "Control_DB".LCnv_Sys[2].Cnv_Level[6].Cnv1.Inputs.Sdetect1 := NOT "C2106 - SHUTTLE IN POSITION 1";
               "Control_DB".LCnv_Sys[2].Cnv_Level[6].Cnv1.Inputs.Sdetect2 := NOT "C2106 - SHUTTLE IN POSITION 2";
               "Control_DB".LCnv_Sys[2].Cnv_Level[6].Cnv1.Safety_Stop_Cnrl.Inputs.DP_Extended := "C2106 - SENSOR SAFETY PIN1 UP";
               "Control_DB".LCnv_Sys[2].Cnv_Level[6].Cnv1.Safety_Stop_Cnrl.Inputs.DP_Retracted := "C2106 - SENSOR SAFETY PIN1 DOWN";

               "Control_DB".LCnv_Sys[2].Cnv_Level[6].Cnv1.Inputs.VFD_Status := "C2106_StatusWord";
               "Control_DB".LCnv_Sys[2].Cnv_Level[6].Cnv1.Inputs.VFD_ActualCurrent := WORD_TO_INT("C2106_ActualCurrent");
               "Control_DB".LCnv_Sys[2].Cnv_Level[6].Cnv1.Inputs.VFD_Speed_Actual := WORD_TO_INT("C2106_ActualSpeed");
               "Control_DB".LCnv_Sys[2].Cnv_Level[6].Cnv1.Inputs.VFD_ActualTorque := WORD_TO_INT("C2106_ActualTorque");

               //BUFFER CONVEYOR LEVEL 6 - CONVEYOR 2
               "Control_DB".LCnv_Sys[2].Cnv_Level[6].Cnv2.Inputs.Left := NOT "C2206 - SENSOR CNV LEFT";
               "Control_DB".LCnv_Sys[2].Cnv_Level[6].Cnv2.Inputs.Lpd1 := NOT "C2206 - SENSOR CNV LEFT (PALLET DETECT 1)";
               "Control_DB".LCnv_Sys[2].Cnv_Level[6].Cnv2.Inputs.Lpd2 := NOT "C2206 - SENSOR CNV LEFT (PALLET DETECT 2)";
               "Control_DB".LCnv_Sys[2].Cnv_Level[6].Cnv2.Inputs.Right := NOT "C2206 - SENSOR CNV RIGHT";
               "Control_DB".LCnv_Sys[2].Cnv_Level[6].Cnv2.Inputs.Rpd1 := NOT "C2206 - SENSOR CNV RIGHT (PALLET DETECT 1)";
               "Control_DB".LCnv_Sys[2].Cnv_Level[6].Cnv2.Inputs.Rpd2 := NOT "C2206 - SENSOR CNV RIGHT (PALLET DETECT 2)";
               "Control_DB".LCnv_Sys[2].Cnv_Level[6].Cnv2.Inputs.Sdetect1 := NOT "C2206 - SHUTTLE IN POSITION 1";
               "Control_DB".LCnv_Sys[2].Cnv_Level[6].Cnv2.Inputs.Sdetect2 := NOT "C2206 - SHUTTLE IN POSITION 2";
               "Control_DB".LCnv_Sys[2].Cnv_Level[6].Cnv2.Safety_Stop_Cnrl.Inputs.DP_Extended := "C2206 - SENSOR SAFETY PIN1 UP";
               "Control_DB".LCnv_Sys[2].Cnv_Level[6].Cnv2.Safety_Stop_Cnrl.Inputs.DP_Retracted := "C2206 - SENSOR SAFETY PIN1 DOWN";

               "Control_DB".LCnv_Sys[2].Cnv_Level[6].Cnv2.Inputs.VFD_Status := "C2206_StatusWord";
               "Control_DB".LCnv_Sys[2].Cnv_Level[6].Cnv2.Inputs.VFD_ActualCurrent := WORD_TO_INT("C2206_ActualCurrent");
               "Control_DB".LCnv_Sys[2].Cnv_Level[6].Cnv2.Inputs.VFD_Speed_Actual := WORD_TO_INT("C2206_ActualSpeed");
               "Control_DB".LCnv_Sys[2].Cnv_Level[6].Cnv2.Inputs.VFD_ActualTorque := WORD_TO_INT("C2206_ActualTorque");
           END_REGION

           REGION LEVEL 7
               //BUFFER CONVEYOR LEVEL 7 - CONVEYOR 1
               "Control_DB".LCnv_Sys[2].Cnv_Level[7].Cnv1.Inputs.Left := NOT "C2107 - SENSOR CNV LEFT";
               "Control_DB".LCnv_Sys[2].Cnv_Level[7].Cnv1.Inputs.Lpd1 := NOT "C2107 - SENSOR CNV LEFT (PALLET DETECT 1)";
               "Control_DB".LCnv_Sys[2].Cnv_Level[7].Cnv1.Inputs.Lpd2 := NOT "C2107 - SENSOR CNV LEFT (PALLET DETECT 2)";
               "Control_DB".LCnv_Sys[2].Cnv_Level[7].Cnv1.Inputs.Right := NOT "C2107 - SENSOR CNV RIGHT";
               "Control_DB".LCnv_Sys[2].Cnv_Level[7].Cnv1.Inputs.Rpd1 := NOT "C2107 - SENSOR CNV RIGHT (PALLET DETECT 1)";
               "Control_DB".LCnv_Sys[2].Cnv_Level[7].Cnv1.Inputs.Rpd2 := NOT "C2107 - SENSOR CNV RIGHT (PALLET DETECT 2)";
               "Control_DB".LCnv_Sys[2].Cnv_Level[7].Cnv1.Inputs.Sdetect1 := NOT "C2107 - SHUTTLE IN POSITION 1";
               "Control_DB".LCnv_Sys[2].Cnv_Level[7].Cnv1.Inputs.Sdetect2 := NOT "C2107 - SHUTTLE IN POSITION 2";
               "Control_DB".LCnv_Sys[2].Cnv_Level[7].Cnv1.Safety_Stop_Cnrl.Inputs.DP_Extended := "C2107 - SENSOR SAFETY PIN1 UP";
               "Control_DB".LCnv_Sys[2].Cnv_Level[7].Cnv1.Safety_Stop_Cnrl.Inputs.DP_Retracted := "C2107 - SENSOR SAFETY PIN1 DOWN";

               "Control_DB".LCnv_Sys[2].Cnv_Level[7].Cnv1.Inputs.VFD_Status := "C2107_StatusWord";
               "Control_DB".LCnv_Sys[2].Cnv_Level[7].Cnv1.Inputs.VFD_ActualCurrent := WORD_TO_INT("C2107_ActualCurrent");
               "Control_DB".LCnv_Sys[2].Cnv_Level[7].Cnv1.Inputs.VFD_Speed_Actual := WORD_TO_INT("C2107_ActualSpeed");
               "Control_DB".LCnv_Sys[2].Cnv_Level[7].Cnv1.Inputs.VFD_ActualTorque := WORD_TO_INT("C2107_ActualTorque");

               //BUFFER CONVEYOR LEVEL 7 - CONVEYOR 2
               "Control_DB".LCnv_Sys[2].Cnv_Level[7].Cnv2.Inputs.Left := NOT "C2207 - SENSOR CNV LEFT";
               "Control_DB".LCnv_Sys[2].Cnv_Level[7].Cnv2.Inputs.Lpd1 := NOT "C2207 - SENSOR CNV LEFT (PALLET DETECT 1)";
               "Control_DB".LCnv_Sys[2].Cnv_Level[7].Cnv2.Inputs.Lpd2 := NOT "C2207 - SENSOR CNV LEFT (PALLET DETECT 2)";
               "Control_DB".LCnv_Sys[2].Cnv_Level[7].Cnv2.Inputs.Right := NOT "C2207 - SENSOR CNV RIGHT";
               "Control_DB".LCnv_Sys[2].Cnv_Level[7].Cnv2.Inputs.Rpd1 := NOT "C2207 - SENSOR CNV RIGHT (PALLET DETECT 1)";
               "Control_DB".LCnv_Sys[2].Cnv_Level[7].Cnv2.Inputs.Rpd2 := NOT "C2207 - SENSOR CNV RIGHT (PALLET DETECT 2)";
               "Control_DB".LCnv_Sys[2].Cnv_Level[7].Cnv2.Inputs.Sdetect1 := NOT "C2207 - SHUTTLE IN POSITION 1";
               "Control_DB".LCnv_Sys[2].Cnv_Level[7].Cnv2.Inputs.Sdetect2 := NOT "C2207 - SHUTTLE IN POSITION 2";
               "Control_DB".LCnv_Sys[2].Cnv_Level[7].Cnv2.Safety_Stop_Cnrl.Inputs.DP_Extended := "C2207 - SENSOR SAFETY PIN1 UP";
               "Control_DB".LCnv_Sys[2].Cnv_Level[7].Cnv2.Safety_Stop_Cnrl.Inputs.DP_Retracted := "C2207 - SENSOR SAFETY PIN1 DOWN";

               "Control_DB".LCnv_Sys[2].Cnv_Level[7].Cnv2.Inputs.VFD_Status := "C2207_StatusWord";
               "Control_DB".LCnv_Sys[2].Cnv_Level[7].Cnv2.Inputs.VFD_ActualCurrent := WORD_TO_INT("C2207_ActualCurrent");
               "Control_DB".LCnv_Sys[2].Cnv_Level[7].Cnv2.Inputs.VFD_Speed_Actual := WORD_TO_INT("C2207_ActualSpeed");
               "Control_DB".LCnv_Sys[2].Cnv_Level[7].Cnv2.Inputs.VFD_ActualTorque := WORD_TO_INT("C2207_ActualTorque");
           END_REGION

           REGION LEVEL 8
               //BUFFER CONVEYOR LEVEL 8 - CONVEYOR 1
               "Control_DB".LCnv_Sys[2].Cnv_Level[8].Cnv1.Inputs.Left := NOT "C2108 - SENSOR CNV LEFT";
               "Control_DB".LCnv_Sys[2].Cnv_Level[8].Cnv1.Inputs.Lpd1 := NOT "C2108 - SENSOR CNV LEFT (PALLET DETECT 1)";
               "Control_DB".LCnv_Sys[2].Cnv_Level[8].Cnv1.Inputs.Lpd2 := NOT "C2108 - SENSOR CNV LEFT (PALLET DETECT 2)";
               "Control_DB".LCnv_Sys[2].Cnv_Level[8].Cnv1.Inputs.Right := NOT "C2108 - SENSOR CNV RIGHT";
               "Control_DB".LCnv_Sys[2].Cnv_Level[8].Cnv1.Inputs.Rpd1 := NOT "C2108 - SENSOR CNV RIGHT (PALLET DETECT 1)";
               "Control_DB".LCnv_Sys[2].Cnv_Level[8].Cnv1.Inputs.Rpd2 := NOT "C2108 - SENSOR CNV RIGHT (PALLET DETECT 2)";
               "Control_DB".LCnv_Sys[2].Cnv_Level[8].Cnv1.Inputs.Sdetect1 := NOT "C2108 - SHUTTLE IN POSITION 1";
               "Control_DB".LCnv_Sys[2].Cnv_Level[8].Cnv1.Inputs.Sdetect2 := NOT "C2108 - SHUTTLE IN POSITION 2";
               "Control_DB".LCnv_Sys[2].Cnv_Level[8].Cnv1.Safety_Stop_Cnrl.Inputs.DP_Extended := "C2108 - SENSOR SAFETY PIN1 UP";
               "Control_DB".LCnv_Sys[2].Cnv_Level[8].Cnv1.Safety_Stop_Cnrl.Inputs.DP_Retracted := "C2108 - SENSOR SAFETY PIN1 DOWN";

               "Control_DB".LCnv_Sys[2].Cnv_Level[8].Cnv1.Inputs.VFD_Status := "C2108_StatusWord";
               "Control_DB".LCnv_Sys[2].Cnv_Level[8].Cnv1.Inputs.VFD_ActualCurrent := WORD_TO_INT("C2108_ActualCurrent");
               "Control_DB".LCnv_Sys[2].Cnv_Level[8].Cnv1.Inputs.VFD_Speed_Actual := WORD_TO_INT("C2108_ActualSpeed");
               "Control_DB".LCnv_Sys[2].Cnv_Level[8].Cnv1.Inputs.VFD_ActualTorque := WORD_TO_INT("C2108_ActualTorque");

               //BUFFER CONVEYOR LEVEL 8 - CONVEYOR 2
               "Control_DB".LCnv_Sys[2].Cnv_Level[8].Cnv2.Inputs.Left := NOT "C2208 - SENSOR CNV LEFT";
               "Control_DB".LCnv_Sys[2].Cnv_Level[8].Cnv2.Inputs.Lpd1 := NOT "C2208 - SENSOR CNV LEFT (PALLET DETECT 1)";
               "Control_DB".LCnv_Sys[2].Cnv_Level[8].Cnv2.Inputs.Lpd2 := NOT "C2208 - SENSOR CNV LEFT (PALLET DETECT 2)";
               "Control_DB".LCnv_Sys[2].Cnv_Level[8].Cnv2.Inputs.Right := NOT "C2208 - SENSOR CNV RIGHT";
               "Control_DB".LCnv_Sys[2].Cnv_Level[8].Cnv2.Inputs.Rpd1 := NOT "C2208 - SENSOR CNV RIGHT (PALLET DETECT 1)";
               "Control_DB".LCnv_Sys[2].Cnv_Level[8].Cnv2.Inputs.Rpd2 := NOT "C2208 - SENSOR CNV RIGHT (PALLET DETECT 2)";
               "Control_DB".LCnv_Sys[2].Cnv_Level[8].Cnv2.Inputs.Sdetect1 := NOT "C2208 - SHUTTLE IN POSITION 1";
               "Control_DB".LCnv_Sys[2].Cnv_Level[8].Cnv2.Inputs.Sdetect2 := NOT "C2208 - SHUTTLE IN POSITION 2";
               "Control_DB".LCnv_Sys[2].Cnv_Level[8].Cnv2.Safety_Stop_Cnrl.Inputs.DP_Extended := "C2208 - SENSOR SAFETY PIN1 UP";
               "Control_DB".LCnv_Sys[2].Cnv_Level[8].Cnv2.Safety_Stop_Cnrl.Inputs.DP_Retracted := "C2208 - SENSOR SAFETY PIN1 DOWN";

               "Control_DB".LCnv_Sys[2].Cnv_Level[8].Cnv2.Inputs.VFD_Status := "C2208_StatusWord";
               "Control_DB".LCnv_Sys[2].Cnv_Level[8].Cnv2.Inputs.VFD_ActualCurrent := WORD_TO_INT("C2208_ActualCurrent");
               "Control_DB".LCnv_Sys[2].Cnv_Level[8].Cnv2.Inputs.VFD_Speed_Actual := WORD_TO_INT("C2208_ActualSpeed");
               "Control_DB".LCnv_Sys[2].Cnv_Level[8].Cnv2.Inputs.VFD_ActualTorque := WORD_TO_INT("C2208_ActualTorque");
           END_REGION
       END_REGION

       REGION VTD
           "Control_DB".VTD_Sys[2].Inputs.Upper_Overtravel :=  "OVERTRAVEL UPPER LIMIT - CH1(2)";
           "Control_DB".VTD_Sys[2].Inputs.Upper_limit := "VTD2 UPPER LIMIT";
           "Control_DB".VTD_Sys[2].Inputs.Ultimate_SlowDown := "VTD2 ULTIMATE SLOWDOWN";
           "Control_DB".VTD_Sys[2].Inputs.Ultimate_Creep := "VTD2 ULTIMATE CREEP";
           "Control_DB".VTD_Sys[2].Inputs.Lower_Limit := "VTD2 LOWER LIMIT";
           "Control_DB".VTD_Sys[2].Inputs.Lower_Overtravel := "OVERTRAVEL LOWER LIMIT - CH1(2)";
           "Control_DB".VTD_Sys[2].Inputs.Level_Detect1 := "VTD2 LEVEL DETECT 1";
           "Control_DB".VTD_Sys[2].Inputs.Level_Detect2 := "VTD2 LEVEL DETECT 2";
           "Control_DB".VTD_Sys[2].Inputs.DP1_Extended := "VTD2 DOCKING PINS EXTENDED 1";
           "Control_DB".VTD_Sys[2].Inputs.DP2_Extended := "VTD2 DOCKING PINS EXTENDED 2";
           "Control_DB".VTD_Sys[2].Inputs.DP1_Retracted := "VTD2 DOCKING PINS RETRACTED 1";
           "Control_DB".VTD_Sys[2].Inputs.DP2_Retracted := "VTD2 DOCKING PINS RETRACTED 2";
           "Control_DB".VTD_Sys[2].Inputs.Chain_Slack_1 := NOT "Remote_Panel_DB_2".Chain_Slack_1_Filtered;
           "Control_DB".VTD_Sys[2].Inputs.Chain_Slack_2 := NOT "Remote_Panel_DB_2".Chain_Slack_2_Filtered;
           "Control_DB".VTD_Sys[2].Inputs.Chain_Slack_3 := NOT "Remote_Panel_DB_2".Chain_Slack_3_Filtered;
           "Control_DB".VTD_Sys[2].Inputs.Chain_Slack_4 := NOT "Remote_Panel_DB_2".Chain_Slack_4_Filtered;
           "Control_DB".VTD_Sys[2].Inputs.PushToEnter := "VTD2 PUSH TO ENTER VTD ZONE";
           "Control_DB".VTD_Sys[2].Inputs.PushToExit := "VTD2 PUSH TO EXIT VTD ZONE";
           "Control_DB".VTD_Sys[2].Inputs.VFD_Status := "VTD2_StatusWord";
           "Control_DB".VTD_Sys[2].Inputs.VFD_ActualCurrent := REAL_TO_INT(("VTD2_ActualCurrent" / 10) / 72.5);
           "Control_DB".VTD_Sys[2].Inputs.VFD_Speed_Actual := "VTD2_ActualSpeed";
           "Control_DB".VTD_Sys[2].Inputs.VFD_ActualTorque := WORD_TO_INT("VTD2_ActualTorque");

       END_REGION

       REGION ABSOLUTE ENCODER
           REGION DOCUMENTATION
               //STATUS---------------------------------------------------------------------------------------------------------------------
               //
               //Encoder state word 2 - INPUT WORD 1
               //
               // 15 … 12 Encoder’s Sign-OF-Life (NOT relevant)
               // 11, 10 Reserved
               // 9 Control requested 0 = No control BY the PLC requested 1 = Control BY the PLC requested
               // 8 … 0 Reserved

               //Sensor 1 state word - INPUT WORD 2
               //
               // 15 Encoder error Description 0 = No error 1 = Error The error code is output in G1_XIST2.
               // 14 Park mode activated 0 = Normal operation 1 = Park mode activated Feedback based on G1_STW bit 14: No output OF position data G1_XIST1 AND G1_XIST2
               // 13 Transmission OF absolute position value 0 = No transmission 1 = Position value is output in G1_XIST2
               // 12 Status OF the Preset function (set/shift OF home position executed) 0 = No Preset function active 1 = Preset function is run Feedback based on G1_STW bit 12:  
               // 11 Requirement OF error acknowledgement detected New position value is output in G1_XIST1 AND G1_XIST2. On conclusion OF the Preset function the bit is set TO 0. 0 = No RETURN acknowledgement OF Encoder error 1 = Requirement OF error acknowledgement detected Reaction TO bit 15 in the sensor control word 1 G1_STW is acknowledged (see Table 14)
               // 10 Reserved
               // 9 … 0 NOT supported

               //Position 1 - INPUT WORD 3 AND 4
               // "AE_Position_1_Scaled" := (*SCALE_X(MIN := "Settings_DB".VTD_Settings.VTD_Min_Height,
               //                                   VALUE := *)NORM_X(MIN := 0,
               //                                                   VALUE := (SHL(IN:="AE_Position_1", N:=2) * 0.00228881) (*- "AE_Offset"*),
               //                                                   MAX := 1073741824)(*,
               //                                   MAX := "Settings_DB".VTD_Settings.VTD_Max_Heigh)*);
               // "mm_per_pulse" := 401,5584 / 262144;
               // 
               //CONTROL---------------------------------------------------------------------------------------------------------------------
               //
               //Encoder control word 2 - OUTPUT WORD 1
               //
               // 15 … 12 Master’s Sign-OF-Life (NOT relevant)
               // 10 control BY PLC 0 = No control BY the PLC 1 = Control BY the PLC Enables the PLC BY using control words TO activate / deactivate encoder functions
               // 7 Fault acknowledge Error-buffer handling NOT supported
               // 11, 9, 8, 6 … 0 Reserved
               // "AE_Control_Word_1".%X10 := "AE_PLC_Control";
               // 
               //Sensor 1 control word - OUTPUT WORD 2-------------------------------------------------------------------------------------------
               //
               // 15 Acknowledging a sensor error Description 0 = Encoder error message NOT acknowledged BY PLC 1 = Encoder error message acknowledged BY the PLC
               // 14 Activate park mode 0 = Normal operation 1 = Activate park mode
               // 13 Request FOR the absolute position value 0 = No request 1 = Request BY the master Results in the cyclic output OF the position values in G1_XIST2
               // 12 Activate preset value (see note below) Defines that a configured preset value is used (see section 3.5 on page 24) 0 = Preset value is NOT activated 1 = Preset value is activated
               // 11 Preset mode Defines how a configured preset value is used 0 = Preset value is used as a new absolute value 1 = Preset value is added TO the previous value
               // 10 … 0 Reserved
               // "AE_Control_Word_2".%X15 := "VTD_Reset_HMI_Tags";
               // "AE_Control_Word_2".%X14 := "AE_Activate_ParkMode";
               // "AE_Control_Word_2".%X13 := "AE_Request_ABS_Value";
               // "AE_Control_Word_2".%X12 := "AE_Activate_Preset_Value";
               // "AE_Control_Word_2".%X11 := "AE_Preset_Mode";
           END_REGION

           //STATUS---------------------------------------------------------------------------------------------------------------------
           "Control_DB".VTD_Sys[2].Inputs.AE_Status_2 := "AE_Status_2(2)";
           //Position 1 - INPUT WORD 3 AND 4
           "Control_DB".VTD_Sys[2].Inputs.AE_Position_1 := REAL_TO_DINT(((((*1073741823 - reverse the direction*)
                                                                                                                                       (SHR(IN := "AE_Position_1(2)", N := 2))) - 31381317) * 0.0015318237304688 (*Mechanical relationship*) + 434391)(*Offset*));

           // Position 2 - INPUT WORD 5 AND 6
           "Control_DB".VTD_Sys[2].Inputs.AE_Position_2 := SHR(IN := "AE_Position_2(2)", N := 2);

           //Speed A - INPUT WORD 7
           "Control_DB".VTD_Sys[2].Inputs.AE_Speed := "AE_Speed(2)";
       END_REGION

       REGION LINEAR ENCODER
           "Control_DB".VTD_Sys[2].Inputs.LE_Position := "LE_X_Unsafe_Position(2)" / 10;
           "Control_DB".VTD_Sys[2].Inputs.LE_Speed := "LE_Speed(2)" * 100;
           "Control_DB".VTD_Sys[2].Inputs.LE_Status := "LE_Status(2)";
           "Control_DB".VTD_Sys[2].Inputs.LE_Warnings := "LE_Warnings(2)";
           REGION DOCUMENTATION
               //STATUS 
               //
               // 0 ERR - Error message (Error code in XP00– XP15); remaining bits = 0, see Error Codes
               // 1 NP - No position information/OUT (XP = 0, YP = 0, SP = 0)
               // 2 WRN - Warnings present, see Warning Module
               // 3 EV - Event present
               // 4 posdetected - Valid position information available

               //WARNINGS
               //
               // 0 WRN01 A code with non-PXV content was found.
               // 1 WRN02 the read head is too close TO the Data Matrix code tape.
               // 2 WRN03 the read head is too far from the Data Matrix code tape.
               // 3 WRN04 Y position too large. The sensor is just before OUT.
               // 4 WRN05 Y position is too small. The sensor is just before OUT.
               // 5 WRN06 the read head is rotated OR tilted in relation TO the Data Matrix code tape.
               // 6 WRN07 Low level OF code contrast.
               // 7 WRN08 Repair tape detected.
               // 8 WRN09 Temperature too high.
               // 9...15 Reserved

               //QUALITY GRADE
               //
               //The quality grades enable constant monitoring of the code tape and the camera along the entire
               //traverse distance. This enables you to detect and act upon potential damage or contamination
               //of the code tape and camera at the earliest stage possible during commissioning and normal
               //operation. As a result, this maximizes the overall functional reliability of your plant, and
               //it means you are able to immediately localize the issue in the case of a fault. Evaluations
               //are made using a scale of 1 to 6. The value 1 is the best possible read quality. A value greater
               //than 3 or worse requires the camera and its path to be inspected. The value 7 signifies "No position"
               //because no code was detected. An evaluation that indicates poor quality as the outcome can be due to
               //a misalignment or incorrect orientation, an incorrect measuring distance, or because the code tape has been affixed incorrectly
           END_REGION
       END_REGION

       REGION SICK BARCODE LECTORS
           IF "Control_DB".VTDBarcode_Station[2].Running AND "SICK_Lector_Control_DB_2".Result <> "Control_DB".VTDBarcode_Station[2].Barcode_Old THEN
               "Control_DB".VTD_Sys[2].Inputs."Barcode 1" := "SICK_Lector_Control_DB_2".Result;
               // "Control_DB".VTD_Control.Inputs."Barcode 2'" := SICK_Barcode_DB".Result;
               // "Control_DB".VTDBarcode_Station[2].Barcode_Old := "SICK_Lector_Control_DB_2".Result;
           ELSE
               "Control_DB".VTD_Sys[2].Inputs."Barcode 1" :=
               "Control_DB".VTD_Sys[2].Inputs."Barcode 2" := '';
           END_IF;

       END_REGION

       REGION VFD HARDWARE ID
           //Buffer conveyors 1
           "Settings_DB".LCnv_Sys[2].Cnv_Level[1].Cnv1.G120_Hardware_ID := "C2101~Drive_1~Standard_telegram_20__PZD-2_6";
           "Settings_DB".LCnv_Sys[2].Cnv_Level[2].Cnv1.G120_Hardware_ID := "C2102~Drive_1~Standard_telegram_20__PZD-2_6";
           "Settings_DB".LCnv_Sys[2].Cnv_Level[3].Cnv1.G120_Hardware_ID := "C2103~Drive_1~Standard_telegram_20__PZD-2_6";
           "Settings_DB".LCnv_Sys[2].Cnv_Level[4].Cnv1.G120_Hardware_ID := "C2104~Drive_1~Standard_telegram_20__PZD-2_6";
           "Settings_DB".LCnv_Sys[2].Cnv_Level[5].Cnv1.G120_Hardware_ID := "C2105~Drive_1~Standard_telegram_20__PZD-2_6";
           "Settings_DB".LCnv_Sys[2].Cnv_Level[6].Cnv1.G120_Hardware_ID := "C2106~Drive_1~Standard_telegram_20__PZD-2_6";
           "Settings_DB".LCnv_Sys[2].Cnv_Level[7].Cnv1.G120_Hardware_ID := "C2107~Drive_1~Standard_telegram_20__PZD-2_6";
           "Settings_DB".LCnv_Sys[2].Cnv_Level[8].Cnv1.G120_Hardware_ID := "C2108~Drive_1~Standard_telegram_20__PZD-2_6";

           //Buffer conveyors 2
           "Settings_DB".LCnv_Sys[2].Cnv_Level[1].Cnv2.G120_Hardware_ID := "C2201~Drive_1~Standard_telegram_20__PZD-2_6";
           "Settings_DB".LCnv_Sys[2].Cnv_Level[2].Cnv2.G120_Hardware_ID := "C2202~Drive_1~Standard_telegram_20__PZD-2_6";
           "Settings_DB".LCnv_Sys[2].Cnv_Level[3].Cnv2.G120_Hardware_ID := "C2203~Drive_1~Standard_telegram_20__PZD-2_6";
           "Settings_DB".LCnv_Sys[2].Cnv_Level[4].Cnv2.G120_Hardware_ID := "C2204~Drive_1~Standard_telegram_20__PZD-2_6";
           "Settings_DB".LCnv_Sys[2].Cnv_Level[5].Cnv2.G120_Hardware_ID := "C2205~Drive_1~Standard_telegram_20__PZD-2_6";
           "Settings_DB".LCnv_Sys[2].Cnv_Level[6].Cnv2.G120_Hardware_ID := "C2206~Drive_1~Standard_telegram_20__PZD-2_6";
           "Settings_DB".LCnv_Sys[2].Cnv_Level[7].Cnv2.G120_Hardware_ID := "C2207~Drive_1~Standard_telegram_20__PZD-2_6";
           "Settings_DB".LCnv_Sys[2].Cnv_Level[8].Cnv2.G120_Hardware_ID := "C2208~Drive_1~Standard_telegram_20__PZD-2_6";

           //Extractor conveyor
           "Settings_DB".ECnv_Sys[2].G120_Hardware_ID := "CVTD_2~Drive_1~Standard_telegram_20__PZD-2_6";

           //VTD
           "Settings_DB".VTD_Sys[2].G120_Hardware_ID := "VTD_2~DO_VECTOR_1~Standard_telegram_20__PZD-2_6";
       END_REGION
   END_REGION

   REGION SYSTEM 3
       REGION EXTRACTOR CONVEYOR
           "Control_DB".ECnv_Sys[3].Inputs.Left := "CVTD3 SENSOR CONVEYOR LEFT (FWD)";
           "Control_DB".ECnv_Sys[3].Inputs.Lpd1 := "CVTD3 SENSOR CONVEYOR LEFT (PALLET DETECT 1)";
           "Control_DB".ECnv_Sys[3].Inputs.Center := "CVTD3 SENSOR CONVEYOR CENTER";
           "Control_DB".ECnv_Sys[3].Inputs.Right := "CVTD3 SENSOR CONVEYOR RIGHT (BWD)";
           "Control_DB".ECnv_Sys[3].Inputs.Rpd1 := "CVTD3 SENSOR CONVEYOR RIGHT (PALLET DETECT 1)";

           "T_OH_Left_3".TOF(IN := "CVTD3 OVERHANG LEFT" OR NOT "Control_DB".VTD_Sys[3].Running,
                             PT := T#200ms);
           "Control_DB".ECnv_Sys[3].Inputs.Overhang_Left := "T_OH_Left_3".Q;

           "T_OH_Right_3".TOF(IN := "CVTD3 OVERHANG RIGHT" OR NOT "Control_DB".VTD_Sys[3].Running,
                              PT := T#200ms);
           "Control_DB".ECnv_Sys[3].Inputs.Overhang_Right := "T_OH_Right_3".Q;

           "Control_DB".ECnv_Sys[3].Inputs.VFD_Status := "CVTD3_StatusWord";
           "Control_DB".ECnv_Sys[3].Inputs.VFD_ActualCurrent := WORD_TO_INT("CVTD3_ActualCurrent");
           "Control_DB".ECnv_Sys[3].Inputs.VFD_Speed_Actual := WORD_TO_INT("CVTD3_ActualSpeed");
           "Control_DB".ECnv_Sys[3].Inputs.VFD_ActualTorque := WORD_TO_INT("CVTD3_ActualTorque");
       END_REGION

       REGION BUFFER CONVEYORS
           REGION LEVEL 1
               //BUFFER CONVEYOR LEVEL 1 - CONVEYOR 1
               "Control_DB".LCnv_Sys[3].Cnv_Level[1].Cnv1.Inputs.Left := NOT "C3101 - SENSOR CNV LEFT (FWD)";
               "Control_DB".LCnv_Sys[3].Cnv_Level[1].Cnv1.Inputs.Lpd1 := NOT "C3101 - SENSOR CNV LEFT (PALLET DETECT 1)";
               "Control_DB".LCnv_Sys[3].Cnv_Level[1].Cnv1.Inputs.Lpd2 := NOT "C3101 - SENSOR CNV LEFT (PALLET DETECT 2)";
               "Control_DB".LCnv_Sys[3].Cnv_Level[1].Cnv1.Inputs.Right := NOT "C3101 - SENSOR CNV RIGHT (BWD)";
               "Control_DB".LCnv_Sys[3].Cnv_Level[1].Cnv1.Inputs.Rpd1 := NOT "C3101 - SENSOR CNV RIGHT (PALLET DETECT 1)";
               "Control_DB".LCnv_Sys[3].Cnv_Level[1].Cnv1.Inputs.Rpd2 := NOT "C3101 - SENSOR CNV RIGHT (PALLET DETECT 2)";
               "Control_DB".LCnv_Sys[3].Cnv_Level[1].Cnv1.Inputs.Sdetect1 := NOT "C3101 - SHUTTLE IN POSITION 1";
               "Control_DB".LCnv_Sys[3].Cnv_Level[1].Cnv1.Inputs.Sdetect2 := NOT "C3101 - SHUTTLE IN POSITION 2";

               "Control_DB".LCnv_Sys[3].Cnv_Level[1].Cnv1.Inputs.VFD_Status := "C3101_StatusWord";
               "Control_DB".LCnv_Sys[3].Cnv_Level[1].Cnv1.Inputs.VFD_ActualCurrent := WORD_TO_INT("C3101_ActualCurrent");
               "Control_DB".LCnv_Sys[3].Cnv_Level[1].Cnv1.Inputs.VFD_Speed_Actual := WORD_TO_INT("C3101_ActualSpeed");
               "Control_DB".LCnv_Sys[3].Cnv_Level[1].Cnv1.Inputs.VFD_ActualTorque := WORD_TO_INT("C3101_ActualTorque");

               //BUFFER CONVEYOR LEVEL 1 - CONVEYOR 2
               "Control_DB".LCnv_Sys[3].Cnv_Level[1].Cnv2.Inputs.Left := NOT "C3201 - SENSOR CNV LEFT (FWD)";
               "Control_DB".LCnv_Sys[3].Cnv_Level[1].Cnv2.Inputs.Lpd1 := NOT "C3201 - SENSOR CNV LEFT (PALLET DETECT 1)";
               "Control_DB".LCnv_Sys[3].Cnv_Level[1].Cnv2.Inputs.Lpd2 := NOT "C3201 - SENSOR CNV LEFT (PALLET DETECT 2)";
               "Control_DB".LCnv_Sys[3].Cnv_Level[1].Cnv2.Inputs.Right := NOT "C3201 - SENSOR CNV RIGHT (BWD)";
               "Control_DB".LCnv_Sys[3].Cnv_Level[1].Cnv2.Inputs.Rpd1 := NOT "C3201 - SENSOR CNV RIGHT (PALLET DETECT 1)";
               "Control_DB".LCnv_Sys[3].Cnv_Level[1].Cnv2.Inputs.Rpd2 := NOT "C3201 - SENSOR CNV RIGHT (PALLET DETECT 2)";
               "Control_DB".LCnv_Sys[3].Cnv_Level[1].Cnv2.Inputs.Sdetect1 := NOT "C3201 - SHUTTLE IN POSITION 1";
               "Control_DB".LCnv_Sys[3].Cnv_Level[1].Cnv2.Inputs.Sdetect2 := NOT "C3201 - SHUTTLE IN POSITION 2";

               "Control_DB".LCnv_Sys[3].Cnv_Level[1].Cnv2.Inputs.VFD_Status := "C3201_StatusWord";
               "Control_DB".LCnv_Sys[3].Cnv_Level[1].Cnv2.Inputs.VFD_ActualCurrent := WORD_TO_INT("C3201_ActualCurrent");
               "Control_DB".LCnv_Sys[3].Cnv_Level[1].Cnv2.Inputs.VFD_Speed_Actual := WORD_TO_INT("C3201_ActualSpeed");
               "Control_DB".LCnv_Sys[3].Cnv_Level[1].Cnv2.Inputs.VFD_ActualTorque := WORD_TO_INT("C3201_ActualTorque");
           END_REGION

           REGION LEVEL 2
               //BUFFER CONVEYOR LEVEL 2 - CONVEYOR 1
               "Control_DB".LCnv_Sys[3].Cnv_Level[2].Cnv1.Inputs.Left := NOT "C3102 - SENSOR CNV LEFT (FWD)";
               "Control_DB".LCnv_Sys[3].Cnv_Level[2].Cnv1.Inputs.Lpd1 := NOT "C3102 - SENSOR CNV LEFT (PALLET DETECT 1)";
               "Control_DB".LCnv_Sys[3].Cnv_Level[2].Cnv1.Inputs.Lpd2 := NOT "C3102 - SENSOR CNV LEFT (PALLET DETECT 2)";
               "Control_DB".LCnv_Sys[3].Cnv_Level[2].Cnv1.Inputs.Right := NOT "C3102 - SENSOR CNV RIGHT (BWD)";
               "Control_DB".LCnv_Sys[3].Cnv_Level[2].Cnv1.Inputs.Rpd1 := NOT "C3102 - SENSOR CNV RIGHT (PALLET DETECT 1)";
               "Control_DB".LCnv_Sys[3].Cnv_Level[2].Cnv1.Inputs.Rpd2 := NOT "C3102 - SENSOR CNV RIGHT (PALLET DETECT 2)";
               "Control_DB".LCnv_Sys[3].Cnv_Level[2].Cnv1.Inputs.Sdetect1 := NOT "C3102 - SHUTTLE IN POSITION 1";
               "Control_DB".LCnv_Sys[3].Cnv_Level[2].Cnv1.Inputs.Sdetect2 := NOT "C3102 - SHUTTLE IN POSITION 2";
               "Control_DB".LCnv_Sys[3].Cnv_Level[2].Cnv1.Safety_Stop_Cnrl.Inputs.DP_Extended := "C3102 - SENSOR SAFETY PIN1 UP";
               "Control_DB".LCnv_Sys[3].Cnv_Level[2].Cnv1.Safety_Stop_Cnrl.Inputs.DP_Retracted := "C3102 - SENSOR SAFETY PIN1 DOWN";

               "Control_DB".LCnv_Sys[3].Cnv_Level[2].Cnv1.Inputs.VFD_Status := "C3102_StatusWord";
               "Control_DB".LCnv_Sys[3].Cnv_Level[2].Cnv1.Inputs.VFD_ActualCurrent := WORD_TO_INT("C3102_ActualCurrent");
               "Control_DB".LCnv_Sys[3].Cnv_Level[2].Cnv1.Inputs.VFD_Speed_Actual := WORD_TO_INT("C3102_ActualSpeed");
               "Control_DB".LCnv_Sys[3].Cnv_Level[2].Cnv1.Inputs.VFD_ActualTorque := WORD_TO_INT("C3102_ActualTorque");

               //BUFFER CONVEYOR LEVEL 2 - CONVEYOR 2
               "Control_DB".LCnv_Sys[3].Cnv_Level[2].Cnv2.Inputs.Left := NOT "C3202 - SENSOR CNV LEFT (FWD)";
               "Control_DB".LCnv_Sys[3].Cnv_Level[2].Cnv2.Inputs.Lpd1 := NOT "C3202 - SENSOR CNV LEFT (PALLET DETECT 1)";
               "Control_DB".LCnv_Sys[3].Cnv_Level[2].Cnv2.Inputs.Lpd2 := NOT "C3202 - SENSOR CNV LEFT (PALLET DETECT 2)";
               "Control_DB".LCnv_Sys[3].Cnv_Level[2].Cnv2.Inputs.Right := NOT "C3202 - SENSOR CNV RIGHT (BWD)";
               "Control_DB".LCnv_Sys[3].Cnv_Level[2].Cnv2.Inputs.Rpd1 := NOT "C3202 - SENSOR CNV RIGHT (PALLET DETECT 1)";
               "Control_DB".LCnv_Sys[3].Cnv_Level[2].Cnv2.Inputs.Rpd2 := NOT "C3202 - SENSOR CNV RIGHT (PALLET DETECT 2)";
               "Control_DB".LCnv_Sys[3].Cnv_Level[2].Cnv2.Inputs.Sdetect1 := NOT "C3202 - SHUTTLE IN POSITION 1";
               "Control_DB".LCnv_Sys[3].Cnv_Level[2].Cnv2.Inputs.Sdetect2 := NOT "C3202 - SHUTTLE IN POSITION 2";
               "Control_DB".LCnv_Sys[3].Cnv_Level[2].Cnv2.Safety_Stop_Cnrl.Inputs.DP_Extended := "C3202 - SENSOR SAFETY PIN1 UP";
               "Control_DB".LCnv_Sys[3].Cnv_Level[2].Cnv2.Safety_Stop_Cnrl.Inputs.DP_Retracted := "C3202 - SENSOR SAFETY PIN1 DOWN";

               "Control_DB".LCnv_Sys[3].Cnv_Level[2].Cnv2.Inputs.VFD_Status := "C3202_StatusWord";
               "Control_DB".LCnv_Sys[3].Cnv_Level[2].Cnv2.Inputs.VFD_ActualCurrent := WORD_TO_INT("C3202_ActualCurrent");
               "Control_DB".LCnv_Sys[3].Cnv_Level[2].Cnv2.Inputs.VFD_Speed_Actual := WORD_TO_INT("C3202_ActualSpeed");
               "Control_DB".LCnv_Sys[3].Cnv_Level[2].Cnv2.Inputs.VFD_ActualTorque := WORD_TO_INT("C3202_ActualTorque");
           END_REGION

           REGION LEVEL 3
               //BUFFER CONVEYOR LEVEL 3 - CONVEYOR 1
               "Control_DB".LCnv_Sys[3].Cnv_Level[3].Cnv1.Inputs.Left := NOT "C3103 - SENSOR CNV LEFT (FWD)";
               "Control_DB".LCnv_Sys[3].Cnv_Level[3].Cnv1.Inputs.Lpd1 := NOT "C3103 - SENSOR CNV LEFT (PALLET DETECT 1)";
               "Control_DB".LCnv_Sys[3].Cnv_Level[3].Cnv1.Inputs.Lpd2 := NOT "C3103 - SENSOR CNV LEFT (PALLET DETECT 2)";
               "Control_DB".LCnv_Sys[3].Cnv_Level[3].Cnv1.Inputs.Right := NOT "C3103 - SENSOR CNV RIGHT (BWD)";
               "Control_DB".LCnv_Sys[3].Cnv_Level[3].Cnv1.Inputs.Rpd1 := NOT "C3103 - SENSOR CNV RIGHT (PALLET DETECT 1)";
               "Control_DB".LCnv_Sys[3].Cnv_Level[3].Cnv1.Inputs.Rpd2 := NOT "C3103 - SENSOR CNV RIGHT (PALLET DETECT 2)";
               "Control_DB".LCnv_Sys[3].Cnv_Level[3].Cnv1.Inputs.Sdetect1 := NOT "C3103 - SHUTTLE IN POSITION 1";
               "Control_DB".LCnv_Sys[3].Cnv_Level[3].Cnv1.Inputs.Sdetect2 := NOT "C3103 - SHUTTLE IN POSITION 2";
               "Control_DB".LCnv_Sys[3].Cnv_Level[3].Cnv1.Safety_Stop_Cnrl.Inputs.DP_Extended := "C3103 - SENSOR SAFETY PIN1 UP";
               "Control_DB".LCnv_Sys[3].Cnv_Level[3].Cnv1.Safety_Stop_Cnrl.Inputs.DP_Retracted := "C3103 - SENSOR SAFETY PIN1 DOWN";

               "Control_DB".LCnv_Sys[3].Cnv_Level[3].Cnv1.Inputs.VFD_Status := "C3103_StatusWord";
               "Control_DB".LCnv_Sys[3].Cnv_Level[3].Cnv1.Inputs.VFD_ActualCurrent := WORD_TO_INT("C3103_ActualCurrent");
               "Control_DB".LCnv_Sys[3].Cnv_Level[3].Cnv1.Inputs.VFD_Speed_Actual := WORD_TO_INT("C3103_ActualSpeed");
               "Control_DB".LCnv_Sys[3].Cnv_Level[3].Cnv1.Inputs.VFD_ActualTorque := WORD_TO_INT("C3103_ActualTorque");

               //BUFFER CONVEYOR LEVEL 3 - CONVEYOR 2
               "Control_DB".LCnv_Sys[3].Cnv_Level[3].Cnv2.Inputs.Left := NOT "C3203 - SENSOR CNV LEFT (FWD)";
               "Control_DB".LCnv_Sys[3].Cnv_Level[3].Cnv2.Inputs.Lpd1 := NOT "C3203 - SENSOR CNV LEFT (PALLET DETECT 1)";
               "Control_DB".LCnv_Sys[3].Cnv_Level[3].Cnv2.Inputs.Lpd2 := NOT "C3203 - SENSOR CNV LEFT (PALLET DETECT 2)";
               "Control_DB".LCnv_Sys[3].Cnv_Level[3].Cnv2.Inputs.Right := NOT "C3203 - SENSOR CNV RIGHT (BWD)";
               "Control_DB".LCnv_Sys[3].Cnv_Level[3].Cnv2.Inputs.Rpd1 := NOT "C3203 - SENSOR CNV RIGHT (PALLET DETECT 1)";
               "Control_DB".LCnv_Sys[3].Cnv_Level[3].Cnv2.Inputs.Rpd2 := NOT "C3203 - SENSOR CNV RIGHT (PALLET DETECT 2)";
               "Control_DB".LCnv_Sys[3].Cnv_Level[3].Cnv2.Inputs.Sdetect1 := NOT "C3203 - SHUTTLE IN POSITION 1";
               "Control_DB".LCnv_Sys[3].Cnv_Level[3].Cnv2.Inputs.Sdetect2 := NOT "C3203 - SHUTTLE IN POSITION 2";
               "Control_DB".LCnv_Sys[3].Cnv_Level[3].Cnv2.Safety_Stop_Cnrl.Inputs.DP_Extended := "C3203 - SENSOR SAFETY PIN1 UP";
               "Control_DB".LCnv_Sys[3].Cnv_Level[3].Cnv2.Safety_Stop_Cnrl.Inputs.DP_Retracted := "C3203 - SENSOR SAFETY PIN1 DOWN";

               "Control_DB".LCnv_Sys[3].Cnv_Level[3].Cnv2.Inputs.VFD_Status := "C3203_StatusWord";
               "Control_DB".LCnv_Sys[3].Cnv_Level[3].Cnv2.Inputs.VFD_ActualCurrent := WORD_TO_INT("C3203_ActualCurrent");
               "Control_DB".LCnv_Sys[3].Cnv_Level[3].Cnv2.Inputs.VFD_Speed_Actual := WORD_TO_INT("C3203_ActualSpeed");
               "Control_DB".LCnv_Sys[3].Cnv_Level[3].Cnv2.Inputs.VFD_ActualTorque := WORD_TO_INT("C3203_ActualTorque");
           END_REGION

           REGION LEVEL 4
               //BUFFER CONVEYOR LEVEL 4 - CONVEYOR 1
               "Control_DB".LCnv_Sys[3].Cnv_Level[4].Cnv1.Inputs.Left := NOT "C3104 - SENSOR CNV LEFT (FWD)";
               "Control_DB".LCnv_Sys[3].Cnv_Level[4].Cnv1.Inputs.Lpd1 := NOT "C3104 - SENSOR CNV LEFT (PALLET DETECT 1)";
               "Control_DB".LCnv_Sys[3].Cnv_Level[4].Cnv1.Inputs.Lpd2 := NOT "C3104 - SENSOR CNV LEFT (PALLET DETECT 2)";
               "Control_DB".LCnv_Sys[3].Cnv_Level[4].Cnv1.Inputs.Right := NOT "C3104 - SENSOR CNV RIGHT (BWD)";
               "Control_DB".LCnv_Sys[3].Cnv_Level[4].Cnv1.Inputs.Rpd1 := NOT "C3104 - SENSOR CNV RIGHT (PALLET DETECT 1)";
               "Control_DB".LCnv_Sys[3].Cnv_Level[4].Cnv1.Inputs.Rpd2 := NOT "C3104 - SENSOR CNV RIGHT (PALLET DETECT 2)";
               "Control_DB".LCnv_Sys[3].Cnv_Level[4].Cnv1.Inputs.Sdetect1 := NOT "C3104 - SHUTTLE IN POSITION 1";
               "Control_DB".LCnv_Sys[3].Cnv_Level[4].Cnv1.Inputs.Sdetect2 := NOT "C3104 - SHUTTLE IN POSITION 2";
               "Control_DB".LCnv_Sys[3].Cnv_Level[4].Cnv1.Safety_Stop_Cnrl.Inputs.DP_Extended := "C3104 - SENSOR SAFETY PIN1 UP";
               "Control_DB".LCnv_Sys[3].Cnv_Level[4].Cnv1.Safety_Stop_Cnrl.Inputs.DP_Retracted := "C3104 - SENSOR SAFETY PIN1 DOWN";

               "Control_DB".LCnv_Sys[3].Cnv_Level[4].Cnv1.Inputs.VFD_Status := "C3104_StatusWord";
               "Control_DB".LCnv_Sys[3].Cnv_Level[4].Cnv1.Inputs.VFD_ActualCurrent := WORD_TO_INT("C3104_ActualCurrent");
               "Control_DB".LCnv_Sys[3].Cnv_Level[4].Cnv1.Inputs.VFD_Speed_Actual := WORD_TO_INT("C3104_ActualSpeed");
               "Control_DB".LCnv_Sys[3].Cnv_Level[4].Cnv1.Inputs.VFD_ActualTorque := WORD_TO_INT("C3104_ActualTorque");

               //BUFFER CONVEYOR LEVEL 4 - CONVEYOR 2
               "Control_DB".LCnv_Sys[3].Cnv_Level[4].Cnv2.Inputs.Left := NOT "C3204 - SENSOR CNV LEFT (FWD)";
               "Control_DB".LCnv_Sys[3].Cnv_Level[4].Cnv2.Inputs.Lpd1 := NOT "C3204 - SENSOR CNV LEFT (PALLET DETECT 1)";
               "Control_DB".LCnv_Sys[3].Cnv_Level[4].Cnv2.Inputs.Lpd2 := NOT "C3204 - SENSOR CNV LEFT (PALLET DETECT 2)";
               "Control_DB".LCnv_Sys[3].Cnv_Level[4].Cnv2.Inputs.Right := NOT "C3204 - SENSOR CNV RIGHT (BWD)";
               "Control_DB".LCnv_Sys[3].Cnv_Level[4].Cnv2.Inputs.Rpd1 := NOT "C3204 - SENSOR CNV RIGHT (PALLET DETECT 1)";
               "Control_DB".LCnv_Sys[3].Cnv_Level[4].Cnv2.Inputs.Rpd2 := NOT "C3204 - SENSOR CNV RIGHT (PALLET DETECT 2)";
               "Control_DB".LCnv_Sys[3].Cnv_Level[4].Cnv2.Inputs.Sdetect1 := NOT "C3204 - SHUTTLE IN POSITION 1";
               "Control_DB".LCnv_Sys[3].Cnv_Level[4].Cnv2.Inputs.Sdetect2 := NOT "C3204 - SHUTTLE IN POSITION 2";
               "Control_DB".LCnv_Sys[3].Cnv_Level[4].Cnv2.Safety_Stop_Cnrl.Inputs.DP_Extended := "C3204 - SENSOR SAFETY PIN1 UP";
               "Control_DB".LCnv_Sys[3].Cnv_Level[4].Cnv2.Safety_Stop_Cnrl.Inputs.DP_Retracted := "C3204 - SENSOR SAFETY PIN1 DOWN";

